(* IEC 61131-3 sources: traffic-lights/PLC_TrafficLights/Class/SafetyCDIAS_Base (part 5) *)

  // if there is a domain info attached
  if (pNameNewElement^ = '@') & ((pNameNewElement + 1)^ = 'D') then
    // check if it's in the actual domain
    if (pNameNewElement + 3)^ = ':' then
      // 1 digit domain number
      RemoteDomain := (pNameNewElement + 2)^ - '0';
    elsif (pNameNewElement + 4)^ = ':' then
      // 2 digits domain number
      RemoteDomain := ((pNameNewElement + 2)^ - '0') * 10 + (pNameNewElement + 3)^ - '0';
    else
      LogError("@ZZZZ (SafetyCDIAS_Base::AddUnsafeRoutElement) Invalid domain info at unsafe variable");
      return;
    end_if;

    // prepare the string (remove the domain info)
    if RemoteDomain >= 10 then
      ui_NameLen      -= 5;
      pNameNewElement += 5;
    else
      ui_NameLen      -= 4;
      pNameNewElement += 4;
    end_if;
  end_if;

  //With the first element, the table must be positioned
  if ( pRoutTable^ = NIL ) then

    //allocate memory for first routing element
    pRoutTable^$^void := To_StdLib.Malloc(size := sizeof(UnsafeIORoutingElement));

    if ( pRoutTable^ = NIL ) then

      State.uiIO_Flags                  := 0;
      State.uiIO_Flags.PhysicAccessOff 	:= 1;
      sd_retval                         :=-1;
      ClassState                        := _MemAllocFailed;
      return;

    end_if;

    p_RoutElement := pRoutTable^;

  else

    //add new element

    //add space for one element to table (linked list element for inputs and linear data area for outputs)
    if LinearMemory = FALSE then
    // search for a place
      p_RoutElement := pRoutTable^;
      while p_RoutElement^.pNext do
        p_RoutElement := p_RoutElement^.pNext;
      end_while;
      p_RoutElement^.pNext$^void := To_StdLib.Malloc(sizeof(UnsafeIORoutingElement));

      if ( p_RoutElement^.pNext = NIL ) then

        State.uiIO_Flags                  := 0;
        State.uiIO_Flags.PhysicAccessOff 	:= 1;
        sd_retval                         :=-1;
        ClassState                        := _MemAllocFailed;
        return;

      end_if;

      // set pointer to new element
      p_RoutElement := p_RoutElement^.pNext;
    else
      pRoutTable^$^void := To_StdLib.ReAlloc(mptr := pRoutTable^, newsize := ( ( pRoutElementsNo^ + 1 ) * sizeof(UnsafeIORoutingElement)));

      if ( pRoutTable^ = NIL ) then

        State.uiIO_Flags                  := 0;
        State.uiIO_Flags.PhysicAccessOff 	:= 1;
        sd_retval                         :=-1;
        ClassState                        := _MemAllocFailed;
        return;

      end_if;

      //set pointer to empty element on last position
      p_RoutElement := pRoutTable^ + ( pRoutElementsNo^ ) * sizeof(UnsafeIORoutingElement);
    end_if;
  end_if;

  if p_RoutElement then
    //allocate memory for name
    p_RoutElement^.pName$^void := To_StdLib.Malloc(size := ui_NameLen);

    if ( p_RoutElement^.pName = NIL ) then

      State.uiIO_Flags                  := 0;
      State.uiIO_Flags.PhysicAccessOff 	:= 1;
      sd_retval                         :=-1;
      ClassState                        := _MemAllocFailed;
      return;

    end_if;

    p_RoutElement^.NameLength := ui_NameLen;
    _memcpy(ptr1:=p_RoutElement^.pName, ptr2:=pNameNewElement, cntr:=ui_NameLen);

    // unsafe bdint variables are localized in a different memory area
    if BitMask then
      p_RoutElement^.ud_Address         := SDO_ADDRESS_UNSAFE_BDINT + ud_Address;
    else
      p_RoutElement^.ud_Address         := SDO_ADDRESS_APP_DATA + ud_Address;
    end_if;

    p_RoutElement^.BitMask              := BitMask;

    // initialize with invalid
    p_RoutElement^.b_IsValid            := FALSE;
    p_RoutElement^.sd_OldValue          := (16#80000000)$DINT;
    p_RoutElement^.sd_NewValue4External := (16#80000000)$DINT;

    // remember that we haven't transmitted this value so far
    p_RoutElement^.b_AlreadyTransmitted := FALSE;

    // initialize next pointer
    p_RoutElement^.pNext                := NIL;

    //increase counter
    pRoutElementsNo^                    += 1;

    // check if name exists in PLC
    p_RoutElement^.ud_Thisp             := GetThisViaServerName(pNameNewElement)$UDINT;
    if (pRoutTable = #p_UnsafeOutputsTable) & p_RoutElement^.BitMask then
      p_RoutElement^.UnsafeType         := BDINTOutput;
    else
      p_RoutElement^.UnsafeType         := NormalUnsafe;
    end_if;
  end_if;

END_FUNCTION

FUNCTION VIRTUAL SafetyCDIAS_Base::InitPathInfo
	VAR_INPUT
		pPathInfo 	: ^PathInfoType;
	END_VAR

  pPathInfo^.p_us_Path      := NIL;
  pPathInfo^.p_us_PathComp  := NIL;
  pPathInfo^.ui_PathCompLen := 0;

END_FUNCTION

FUNCTION VIRTUAL SafetyCDIAS_Base::WriteTDO2Module
	VAR_INPUT
		pTDO 	: ^TDOType;
	END_VAR
#ifdef SAFETY_OVER_DIAS
  VAR
    i : DINT;
  END_VAR
#endif

  if ( State.uiIO_Flags = 0 ) then

  #ifdef SAFETY_OVER_DIAS
    #pragma message("TDO-Handling over DIAS has to be reworked!")
    if ( b_im ) then
      //copy TDO word by word
      for i := 0 to (((TDOInfo AND 16#7F)/2)-1) by 1 do

        ( a_Handle_TDO_Write[i] )$^UINT^ := ( (pTDO)$^UINT + ( i * 2 ) )^;

      end_for;
    else
  #endif

      // responses into response buffer, request into requestbuffer (only enough place for 1)
      if pTDO^.StdHeader.Typ AND SSDO_MASK_RESPONSE then
        IF ( s_TDORingbuffer.ud_entries < ( SIZEOF( TDORingbuffer.Entry ) / SIZEOF( TDOType ) ) ) THEN
          s_TDORingbuffer.Entry[s_TDORingbuffer.ud_WritePos] :=  pTDO^;
          s_TDORingbuffer.ud_WritePos       := ( s_TDORingbuffer.ud_WritePos + 1 ) mod ( SIZEOF( TDORingbuffer.Entry ) / SIZEOF( TDOType ) );
          s_TDORingbuffer.ud_Entries        += 1;
          s_TDORingbuffer.b_ErrorTriggered  := FALSE;
        ELSIF ( s_TDORingbuffer.b_ErrorTriggered = FALSE ) THEN
          LogError("@ZZZZ (SafetyCDIAS_Base::WriteTDO2Module) [SL] Buffer for TDO-Messages is full!");
          s_TDORingbuffer.b_ErrorTriggered  := TRUE;
        END_IF;

        IF s_TDORingbuffer.ud_Entries > s_TDORingbuffer.ud_maxEntries THEN
          s_TDORingbuffer.ud_maxEntries     := s_TDORingbuffer.ud_Entries;
        END_IF;
      else
        s_TDORingbuffer.RequestTDO          := pTDO^;
        s_TDORingbuffer.b_RequestAvailable  := TRUE;
      end_if;

  #ifdef SAFETY_OVER_DIAS
    end_if;
  #endif
  end_if;

END_FUNCTION

FUNCTION VIRTUAL SafetyCDIAS_Base::ResetConfig
  VAR
    p_SafetyBase        : pVirtualBase;
  	p_RoutElement       : ^RoutElement;
    p_UnsafeRoutElement : ^UnsafeIORoutingElement;
    i                   : UINT;
    ii                  : DINT;
		MyPara 	            : CmdStruct;
		MyResult	          : results;
  END_VAR

  // tell all modules, which are connected to this cpu (through the old configuration) that they should delete the cpu from their routing table
  // must be more than 1, because 1st is always own entry
  if p_RoutTable & (ui_CntRoutElements > 1) then
    //set pointer on 2nd routing element
    p_RoutElement := p_RoutTable + sizeof(RoutElement);
    for i := 1 to (ui_CntRoutElements - 1) do
      // clear everything except this object (done after the for loop)
      if p_RoutElement^.ud_Thisp <> THIS$UDINT then
        // get thispointer of routing element
        p_SafetyBase := (p_RoutElement^.ud_Thisp)$pVirtualBase;

        // call other safety-class to remove the safetynumber from the routing table
        MyPara.uiCmd := CMD_SM_REMOVE_CPU_FROM_TABLE;
        MyPara.aPara[0] := SafetyNumber$DINT;

        p_SafetyBase^.NewInst(#MyPara, #MyResult);

//        p_SafetyBase^.RemoveCPUFromTable(ud_SafetyNr := SafetyNumber);
      end_if;

      // free memory of compressed path
      if p_RoutElement^.p_CompressedPath then
        To_StdLib.Free(mptr:=p_RoutElement^.p_CompressedPath);
      end_if;

      // set pointer on next routing element
      p_RoutElement += sizeof(RoutElement);
    end_for;

    // reduce local routing table to the cpu's own entry
    ui_CntRoutElements := 1;
  end_if;

  // on CSCP011 the SDO_COMMAND_WRITE_VALUES didn't exist, so we have to make a difference here
  if (us_Variant <> CSCP011_Preliminary) & (us_Variant <> CSCP011_Preliminary) then
    while p_UnsafeInputsTable do
      p_UnsafeRoutElement := p_UnsafeInputsTable;
      p_UnsafeInputsTable := p_UnsafeInputsTable^.pNext;

      To_StdLib.Free(mptr:=p_UnsafeRoutElement^.pName);
      To_StdLib.Free(mptr:=p_UnsafeRoutElement);
    end_while;
  else
    // free list of unsafe elements
    if p_UnsafeInputsTable then
      To_StdLib.Free(mptr:=p_UnsafeInputsTable);
      p_UnsafeInputsTable := NIL;
    end_if;
  end_if;
  ui_CntUnsafeInputs    := 0;

  // unsafe outputs are always in linear memory
  if p_UnsafeOutputsTable then
    To_StdLib.Free(mptr:=p_UnsafeOutputsTable);
    p_UnsafeOutputsTable := NIL;
  end_if;
  ui_CntUnsafeOutputs   := 0;

  // reset no of SDO input buffer
  ui_cnt_SDOInputBuffer := 0;

  // if the old configuration is reset, check for the configured state of the cpu
  b_CheckConfigured     := TRUE;

  if b_VaranAvailable then
    // by default the mover is invalid. it will be initialized when reading the configuration
    b_MoveCommandInputActive  := _Invalid;
    b_MoveCommandOutputActive := _Invalid;

    if b_PayloadSupport then

      DisableDO(ud_DOHandle := InputMovHandle$UDINT);

      if AdditionalSPDOs then
        for ii := 0 to (AdditionalSPDOs-1) do
          DisableDO(ud_DOHandle := aAdditionalPDOs[ii].InputMovHandle$UDINT);
        end_for;
      end_if;
    else

      if InputMovHandle then
        InputMovHandle^.ucCtrlStat := VARAN_DO_NO_RUN;
      end_if;

      if AdditionalSPDOs then
        for ii := 0 to (AdditionalSPDOs-1) do
          aAdditionalPDOs[ii].InputMovHandle^.ucCtrlStat := VARAN_DO_NO_RUN;
        end_for;
      end_if;
    end_if;

  else
    // if no VARAN, we can't move the PDOs
    b_MoveCommandInputActive  := _Inactive;
    b_MoveCommandOutputActive := _Inactive;
  end_if;

END_FUNCTION

FUNCTION VIRTUAL GLOBAL SafetyCDIAS_Base::MyBackground
  VAR
  	sd_retval         : DINT;
    GetStateResp      : GetStateResponseType;
    LastWriteCounter  : UDINT;
    FileHandle        : DINT;
		MyPara 	          : CmdStruct;
		MyResult	        : results;
  END_VAR

  // if any LED is active, then firmware update is not active and we can do our work
  if (VoltageOK | RunState | ServiceMode | Error) then

    // if a quit error is pending
    if QuitComError = 2 then
      MyPara.uiCmd := CMD_SM_QUIT_ERROR_VIA_OS;
      MyPara.aPara[0] := THIS$DINT;
      MyPara.aPara[1] := SafetyNumber$DINT;
      pSafetyManagerThis^.NewInst(#MyPara, #MyResult);

      QuitComError := MyResult.aData[0]$DINT;
    end_if;

    if (ClassState = _ReinitConfig) then

      // check every second if the cpu is configured
      if b_CheckConfigured & ((ops.tAbsolute - ud_LastCheckConfig) > 3000) then
        // get state via SDO communication
        sd_retval := SDOStdRequ ( us_Command      := SDO_COMMAND_GET_STATE
                                , p_us_RespData   := ( #GetStateResp )$^USINT
                                , us_RespLength   := sizeof(GetStateResponseType)
                                );

        // the cpu is configured, load the new configuration
        if ( sd_retval = 0 ) &
           (GetStateResp.ConfigState <> CFG_STATE_UNKNOWN) &
           (GetStateResp.ConfigState <> CFG_STATE_INVALID) &
           (GetStateResp.ConfigState <> CFG_STATE_NOT_CONFIGURED) then

          b_CheckConfigured := FALSE;
          b_GetNewConfiguration := TRUE;
        end_if;

        // remember the last time we checked for configurated cpu
        ud_LastCheckConfig := ops.tAbsolute;
      end_if;

      // if there is a new configuration => get it
      if b_GetNewConfiguration then

        //get configuration from safe CPU and build routing tables
        sd_retval := GetRoutingData();
        if sd_retval = 0 then
          b_GetNewConfiguration := FALSE;

          SendAllUnsafeValues();
        else
          LogError("@ZZZZ (SafetyCDIAS_Base::MyBackground) FAILED TO REINIT THE SAFECPU: ");
        end_if;
      end_if;
    end_if;

    // here we save the log file from the module to the harddrive (started by user)
    if DiagVars.SavingLogInProgress then

      case DiagVars.SavingLogSSW of

  // ********************************************************************************************************************************************
        GetLogHeader:     // get log header from module (contains size of log memory and write counter)

          // get log header via SDO communication
          sd_retval := SDORequ ( us_Command      := SDO_COMMAND_GET_LOG_HDR
                               , p_us_RequData   := #DiagVars.ucChoiceSaveLog
                               , us_RequLength   := 1
                               , p_us_RespData   := ( #DiagVars.LogHeader)$^USINT
                               , us_RespLength   := sizeof(DiagStructType.LogHeader)
                               );

          if ( sd_retval = 0 ) then
            DiagVars.LogMemToGet := DiagVars.LogHeader.LogMemSize;
            DiagVars.pLogFileMem$pVoid := To_StdLib.Malloc(size:=DiagVars.LogHeader.LogMemSize);
            //_memset(dest:=DiagVars.pLogFileMem$pVoid, usByte:=0, cntr:=DiagVars.LogHeader.LogMemSize);
            if DiagVars.ucChoiceSaveLog = 0 then
              DiagVars.ReadBaseAdr  := SDO_ADDRESS_LOG_UC1;
            else
              DiagVars.ReadBaseAdr  := SDO_ADDRESS_LOG_UC2;
            end_if;
            DiagVars.SavingLogSSW   := GetLogFileBlocks;

          end_if;

  // ********************************************************************************************************************************************
        GetLogFileBlocks: // get the log memory from the application memory of the module (every cycle only a little bit to prevent runtime error in module)

          // we wait here until UpdateCy finishes our work

  // ********************************************************************************************************************************************
        GetLogHeader2:    // get log header from module again. if write counter changed,
                          // we repeat GetLogFileBlocks. otherwise we continue to save the file

          LastWriteCounter := DiagVars.LogHeader.WriteCounter;

          // get LogHeader
          sd_retval := SDORequ ( us_Command      := SDO_COMMAND_GET_LOG_HDR
                               , p_us_RequData   := #DiagVars.ucChoiceSaveLog
                               , us_RequLength   := 1
                               , p_us_RespData   := ( #DiagVars.LogHeader)$^USINT
                               , us_RespLength   := sizeof(DiagStructType.LogHeader)
                               );

          if ( sd_retval = 0 ) then

            // if write counter is different, repeat last step
            if DiagVars.LogHeader.WriteCounter <> LastWriteCounter then
              DiagVars.SavingLogSSW := GetLogFileBlocks;

              DiagVars.LogMemToGet := DiagVars.LogHeader.LogMemSize;

              // realloc memory (maybe it's a different size)
              To_StdLib.Free(mptr:=DiagVars.pLogFileMem$pVoid);
              DiagVars.pLogFileMem$pVoid := To_StdLib.Malloc(size:=DiagVars.LogHeader.LogMemSize);
            else
              // write counter is equal. continue to last step
              DiagVars.SavingLogSSW := SaveLogFile;
            end_if;
          end_if;

  // ********************************************************************************************************************************************
        SaveLogFile:      // save the memory to the specified file (DPNE)
          // open file (create/overwrite always)
          FileHandle := FileSys.FileOpen(filename:=#DiagVars.DPNE[0], attributes:=ATT_CREATE_ALWAYS);

          DiagVars.SavingLogSuccessful := 1;

          if FileHandle >= 0 then

            // save content to it
            if FileSys.FileWrite(handle:=FileHandle, buffer:=DiagVars.pLogFileMem, length:=DiagVars.LogHeader.LogMemSize) <> DiagVars.LogHeader.LogMemSize$DINT then
              // failed to write to file
              LogError("@ZZZZ (SafetyCDIAS_Base::MyBackground) Failed to write to binary LogFile");
              DiagVars.SavingLogSuccessful := -1;
            end_if;

            // close file
            FileSys.FileClose(handle:=FileHandle);
          else
            // failed to open file
            LogError("@ZZZZ (SafetyCDIAS_Base::MyBackground) Failed to open binary LogFile");
            DiagVars.SavingLogSuccessful := -1;
          end_if;

          To_StdLib.Free(mptr:=DiagVars.pLogFileMem$pVoid);
          DiagVars.pLogFileMem := NIL;

          DiagVars.SavingLogSSW         := GetLogHeader;
          DiagVars.SavingLogInProgress  := FALSE;

      end_case;
    end_if;
  end_if;

END_FUNCTION

FUNCTION VIRTUAL SafetyCDIAS_Base::RemoveCPUFromTable
	VAR_INPUT
		ud_SafetyNr 	  : HDINT;
	END_VAR
  VAR
  	p_RoutElement   : ^RoutElement;
    i               : UDINT;
    FoundIndex      : UDINT;
    pPDOInputBuffer : ^PDOInputBuffer;
    Found : BOOL;
  END_VAR

  // if we are a cpu, do nothing
  if b_CheckCRC then
    return;
  end_if;

  //check each element (must be more than 1, because 1st is always own entry)
  if p_RoutTable & (ui_CntRoutElements > 1) then
    //set pointer on 2nd routing element
    p_RoutElement := p_RoutTable + sizeof(RoutElement);
    for i := 1 to (ui_CntRoutElements - 1) do

      // if we found safenumber, delete element from table
      if ( p_RoutElement^.ud_SafeNumber = ud_SafetyNr ) then

        // at last element we don't need to copy data, just decrease buffersize
        if i <> (ui_CntRoutElements - 1) then
          _memcpy(p_RoutElement, p_RoutElement + sizeof(RoutElement), sizeof(RoutElement) * (ui_CntRoutElements - 1 - i));
        end_if;

        // free 1 element and decrease element counter
        ui_CntRoutElements -= 1;

        exit;
      end_if;

      // set pointer on next routing element
      p_RoutElement += sizeof(RoutElement);
    end_for;
  end_if;

  // reset no of SDO input buffer
  ui_cnt_SDOInputBuffer := 0;

  if b_VaranAvailable then
    // by default the mover is invalid. it will be initialized when reading the configuration
    b_MoveCommandInputActive  := _Invalid;
    b_MoveCommandOutputActive := _Invalid;

    if InputMovHandle then
      if b_PayloadSupport then
        DisableDO(ud_DOHandle := InputMovHandle$UDINT);

        if AdditionalSPDOs then
          for i := 0 to (AdditionalSPDOs-1)$UDINT do
            DisableDO(ud_DOHandle := aAdditionalPDOs[i].InputMovHandle$UDINT);
          end_for;
        end_if;
      else
        InputMovHandle^.ucCtrlStat := VARAN_DO_NO_RUN;

        if AdditionalSPDOs then
          for i := 0 to (AdditionalSPDOs-1)$UDINT do
            aAdditionalPDOs[i].InputMovHandle^.ucCtrlStat := VARAN_DO_NO_RUN;
          end_for;
        end_if;

      end_if;
    end_if;
  else
    // if no VARAN, we can't move the PDOs
    b_MoveCommandInputActive  := _Inactive;
    b_MoveCommandOutputActive := _Inactive;
  end_if;

  // check if we received a PDO from this CPU => if so, delete it from the PDO input buffer
  if ui_cnt_PDOInputBuffer then
    // search for the PDO
    Found := FALSE;
    pPDOInputBuffer := #aPDOInputBuffer[0];
    for FoundIndex := 0 to (ui_cnt_PDOInputBuffer-1) do
      if pPDOInputBuffer^.ud_SafetyNr = ud_SafetyNr then
        Found := TRUE;
        exit;
      end_if;

      pPDOInputBuffer += sizeof(PDOInputBuffer);
    end_for;

    // if we found the PDO => remove it from memory (move the memory behind the found PDO over the place of the found PDO)
    if Found then
      // if it's last entry (no entries have to be moved) => we only have to copy some memory if it's not the last
      if FoundIndex < (ui_cnt_PDOInputBuffer-1) then
        for i := FoundIndex to (ui_cnt_PDOInputBuffer-2) do
          aPDOInputBuffer[i] := aPDOInputBuffer[i+1];
        end_for;
      end_if;
      ui_cnt_PDOInputBuffer -= 1;
    end_if;
  end_if;

END_FUNCTION

FUNCTION VIRTUAL SafetyCDIAS_Base::CheckUnsafeUpdateCycle

  // we can only use 56 byte pay load (instead of 64) because fw drops the 8 byte used for addresses in safe SDO

  if ui_CntUnsafeOutputs then
  // maximum of read variables in 1 frame is 15 (56 Bytes pay load - 1 Byte Returncode - 1 Byte Length = 54 Bytes => 13x4Bytes = 52)
    MaxVarsPerReadPackage := (SDO_MAX_LENGTH - (sizeof(SDOHeader) - sizeof(SDOHeader.SessId)) - sizeof(SDORespReadConfig.us_Returncode) - sizeof(SDORespReadConfig.us_Length)) / sizeof(DINT);
    ReadFramesNeeded := ((ui_CntUnsafeOutputs - 1) / MaxVarsPerReadPackage) + 1;
  else
    ReadFramesNeeded := 0;
  end_if;

  if ui_CntUnsafeInputs then
  // maximum of write variables in 1 frame is 14 (56 Bytes pay load - 4 Byte Address - 1 Byte Length = 51 Bytes => 12x4Bytes = 48)
    MaxVarsPerWritePackage := (SDO_MAX_LENGTH - (sizeof(SDOHeader) - sizeof(SDOHeader.SessId)) - sizeof(SDORequReadConfig.ud_Address) - sizeof(SDORequReadConfig.us_Length)) / sizeof(DINT);
    WriteFramesNeeded := ((ui_CntUnsafeInputs - 1) / MaxVarsPerWritePackage) + 1;
  else
    WriteFramesNeeded := 0;
  end_if;

  // check if user has given us enough time
  if b_VaranAvailable then
    if sd_VaranType = 2 then
      ud_TransfertimePerPackage := SDO_TRANSFERTIME_MOVER;
    else
      ud_TransfertimePerPackage := SDO_TRANSFERTIME_VARAN;
    end_if;
  else
    ud_TransfertimePerPackage := SDO_TRANSFERTIME_CDIAS;
#ifdef SAFETY_OVER_DIAS
    #pragma message("Transfer time for DIAS must be defined!")
#endif
  end_if;

  if ( (WriteFramesNeeded + ReadFramesNeeded) * ud_TransfertimePerPackage ) > ServerUpdateTime then
    ServerUpdateTime    := ( WriteFramesNeeded + ReadFramesNeeded ) * ud_TransfertimePerPackage;
    ServerUpdateTime.Write(input:=ServerUpdateTime);
    ud_ServerUpdateTime := ( ReadFramesNeeded ) * ud_TransfertimePerPackage;
  end_if;

END_FUNCTION

FUNCTION VIRTUAL GLOBAL SafetyCDIAS_Base::FetchDiagState

  DiagVars.UserDiagStateReady := FALSE;
  DiagVars.UserWantsDiagState := TRUE;

END_FUNCTION

FUNCTION VIRTUAL GLOBAL SafetyCDIAS_Base::GetDiagState
	VAR_INPUT
		pDiagState 	: ^SafetyDiagState;
	END_VAR
	VAR_OUTPUT
		StateReady 	: BOOL;
	END_VAR

  StateReady                        := DiagVars.UserDiagStateReady;

  // if data ready, we save it into user structure
  if StateReady then
    pDiagState^.RunState            := DiagVars.UserGetStateResp.RuntimeState;
    pDiagState^.ConfigState         := DiagVars.UserGetStateResp.ConfigState;
    pDiagState^.LoginLevel          := DiagVars.UserGetStateResp.LoginLevel;
    pDiagState^.ErrorCounterIOState := DiagVars.UserGetStateResp.ErrorCount;
  end_if;

END_FUNCTION

FUNCTION VIRTUAL GLOBAL SafetyCDIAS_Base::FetchDiagInfo
	VAR_INPUT
		ucChoice 	: USINT;
	END_VAR

  DiagVars.ucChoiceDiagInfo  := ucChoice;
  DiagVars.UserDiagInfoReady := FALSE;
  DiagVars.UserWantsDiagInfo := TRUE;

END_FUNCTION

FUNCTION VIRTUAL GLOBAL SafetyCDIAS_Base::GetDiagInfo
	VAR_INPUT
		pDiagInfo 	: ^SafetyDiagInfo;
	END_VAR
	VAR_OUTPUT
		StateReady 	: BOOL;
	END_VAR

  StateReady    := DiagVars.UserDiagInfoReady;

  // if data ready, we save it into user structure
  if StateReady then
    pDiagInfo^  := DiagVars.UserGetDiagInfoResp;
  end_if;

END_FUNCTION

FUNCTION VIRTUAL SafetyCDIAS_Base::SDORequ
	VAR_INPUT
		us_Command 	        : USINT;
		p_us_RequData 	    : ^USINT;
		us_RequLength 	    : USINT;
		p_us_RespData 	    : ^USINT;
		us_RespLength 	    : USINT;
	END_VAR
	VAR_OUTPUT
		sd_retval 	        : DINT;
	END_VAR
  VAR
  	pSDORequestBuffer   : ^SDOStdHeader;
    pSDOResponseBuffer  : ^SDOStdResp;
    RespBuffer          : ARRAY [0..127] OF USINT;
    RequBuffer          : ARRAY [0..127] OF USINT;
    us_InLength         : USINT;
    us_OutLength        : USINT;
  END_VAR

  //SDO requests for this commands don't have any further data
  pSDORequestBuffer$^void   := #RequBuffer[0];
  pSDOResponseBuffer$^void  := #RespBuffer[0];

  //SDO request buffer (length header + data)
  us_InLength               := sizeof(SDOStdHeader) + us_RequLength;

  //SDO response buffer (length header + rc + data)
  us_OutLength              := sizeof(SDOStdHeader) + 1 + us_RespLength;

  //calculate length without crc
  pSDORequestBuffer^.len    := sizeof(SDOStdHeader) - sizeof(SDOStdHeader.CRC) + us_RequLength;

  //type
  pSDORequestBuffer^.typ    := FRM_TYPECODE_STD;

  //sequence number
  pSDORequestBuffer^.SeqNr  := us_CntSequNr;

  _memcpy(ptr1:=pSDORequestBuffer + sizeof(SDOStdHeader), ptr2:=p_us_RequData, cntr:=us_RequLength);

  //increase counter for sequence number
  if us_CntSequNr < 16#7F then
    us_CntSequNr += 1;
  else
    us_CntSequNr := 0;
  end_if;

  //command to inform CPU about initializing classes is ok
  pSDORequestBuffer^.cmd := us_Command;

  //set CRC-field to 0
  pSDORequestBuffer^.CRC := 0;

  //send request
  sd_retval := SAFETY_iSendRequest( uiMaster    := 0
                                  , pucNode     := p_ObjectPath
                                  , uiInLength  := us_InLength
                                  , pucInput    := pSDORequestBuffer$^USINT
                                  , uiOutLength := us_OutLength
                                  , pucOutput   := pSDOResponseBuffer$^USINT
                                  );

  //no response
  if ( sd_retval = 0 ) then

    //check sequence number to exclude a possible wrong response
    if ( pSDORequestBuffer^.SeqNr <> pSDOResponseBuffer^.StdHeader.SeqNr ) then
      sd_retval := -102;

    //check returncode of SDO
    elsif ( pSDOResponseBuffer^.us_Returncode <> SDO_RETCODE_OK ) then
      sd_retval := -103;
    end_if;

  end_if;

  //return response
  if ( ( sd_retval = 0 ) & ( p_us_RespData <> NIL )) then
    To_StdLib.MemCpy(dest := p_us_RespData, source := #pSDOResponseBuffer^.us_Data, size := us_RespLength);
  end_if;

END_FUNCTION

FUNCTION VIRTUAL GLOBAL SafetyCDIAS_Base::SaveLog
	VAR_INPUT
		ucChoice  : USINT;
		pDPNE 	  : ^CHAR;
	END_VAR
	VAR_OUTPUT
		Success 	: DINT;
	END_VAR

  if DiagVars.SavingLogInProgress = FALSE then
    DiagVars.SavingLogInProgress  := TRUE;

    DiagVars.SavingLogSuccessful  := FALSE; //Reset Value

    DiagVars.ucChoiceSaveLog      := ucChoice;

    _memcpy(ptr1:=#DiagVars.DPNE, ptr2:=pDPNE, cntr:=_strlen(pDPNE));

    Success := TRUE;
  else
    Success := FALSE;
  end_if;

END_FUNCTION

FUNCTION VIRTUAL GLOBAL SafetyCDIAS_Base::SaveLogActive
	VAR_OUTPUT
		InProgress 	: BOOL;
	END_VAR

  InProgress := DiagVars.SavingLogInProgress;

END_FUNCTION

FUNCTION VIRTUAL SafetyCDIAS_Base::BlockedTransferLength
	VAR_INPUT
		ud_Datalength 	    : UDINT;
		us_MaxBlocklength 	: USINT;
	END_VAR
	VAR_OUTPUT
		us_ActBlocklength 	: USINT;
	END_VAR

  IF ud_Datalength > to_UDINT(us_MaxBlocklength) THEN
    us_ActBlocklength := us_MaxBlocklength;
  ELSE
    us_ActBlocklength := to_USINT(ud_Datalength);
  END_IF;

END_FUNCTION

FUNCTION VIRTUAL SafetyCDIAS_Base::AddToPDOMoverList
	VAR_INPUT
		pThis 	: pVirtualBase;
		pList 	: ^pPDOMoverList;
	END_VAR
  VAR
    pHelp : ^PDOMoverList;
  END_VAR

  if pList^ = NIL then
    pList$^pvoid^ := To_StdLib.Malloc(size:=sizeof(PDOMoverList));
    //Graphic.Memory((#pList)$^pVoid, sizeof(PDOMoverList));
    pHelp := pList^;
  else
    pHelp := pList^;
    if pHelp^.pThis = pThis then
      // this pointer already in buffer => leave function
      return;
    end_if;
    while pHelp^.pNext <> NIL do
      if pHelp^.pThis <> pThis then
        pHelp := pHelp^.pNext;
      else
        // this pointer already in buffer => leave function
        return;
      end_if;
    end_while;
    pHelp^.pNext$pvoid := To_StdLib.Malloc(size:=sizeof(PDOMoverList));
    pHelp := pHelp^.pNext;
  end_if;

  if pHelp <> NIL then
    pHelp^.pThis := pThis;
    pHelp^.pNext := NIL;
  end_if;

END_FUNCTION

FUNCTION VIRTUAL SafetyCDIAS_Base::WalkThroughPDOMoverList
	VAR_INPUT
		pList 	  : ^pPDOMoverList;
		NewState 	: PDOMoveState;
	END_VAR
  VAR
  	pAct      : ^PDOMoverList;
    pFree     : ^void;
		MyPara 	  : CmdStruct;
		MyResult  : results;
  END_VAR

  // get pointer on first element of list
  pAct := pList^;

  // if we have entries left we walk on
  WHILE pAct DO
#pragma warning(disable:137 )
    // set state of corresponding PDOMover to off
    IF pList = #pPDOMoverListInputs THEN
      if NewState = _Inactive then

        MyPara.uiCmd    := CMD_SM_DEACTIVATE_MOVE_CMD;
        MyPara.aPara[0] := 0;
        pAct^.pThis^.NewInst(#MyPara, #MyResult);

//        pAct^.pThis^.b_MoveCommandOutputActive := _Inactive;
      end_if;
    ELSE
      if NewState = _Inactive then

        MyPara.uiCmd    := CMD_SM_DEACTIVATE_MOVE_CMD;
        MyPara.aPara[0] := 1;
        pAct^.pThis^.NewInst(#MyPara, #MyResult);

//        pAct^.pThis^.b_MoveCommandInputActive := _Inactive;
      end_if;
    END_IF;
#pragma warning(default:137 )

    //go to next entry and get rid of the allocated memory
    pFree := pAct;
    pAct  := pAct^.pNext;
    To_StdLib.Free(mptr:=pFree);
  END_WHILE;

  // we got rid of the memory above - to make sure nobody will use this data again we clear the list entry
  pList^ := NIL;

END_FUNCTION

FUNCTION VIRTUAL SafetyCDIAS_Base::CleanupPDOMoverList
	VAR_INPUT
		pList 	: ^pPDOMoverList;
	END_VAR
  VAR
  	pAct    : ^PDOMoverList;
    pFree   : ^void;
  END_VAR

  // get pointer on first element of list
  pAct := pList^;

  // if we have entries left we walk on
  WHILE pAct DO
    //go to next entry and get rid of the allocated memory
    pFree := pAct;
    pAct  := pAct^.pNext;
    To_StdLib.Free(mptr:=pFree);
  END_WHILE;

  // we got rid of the memory above - to make sure nobody will use this data again we clear the list entry
  pList^ := NIL;

END_FUNCTION

#pragma warning(disable: 73)
FUNCTION VIRTUAL SafetyCDIAS_Base::AddFrame
	VAR_INPUT
		pFrame 	        : ^SafetyCDIAS_Base::SDOStdHeader;
		FrameState 	    : DINT;
		CallerSafetyNr 	: HDINT;
	END_VAR

END_FUNCTION
#pragma warning(default: 73)

FUNCTION VIRTUAL SafetyCDIAS_Base::RecordFrame
	VAR_INPUT
		pFrame 	    : ^DINT;
		FrameState 	: DINT;
	END_VAR
  VAR
    ThisBackup  : pVoid;
    TempSafetyNr: HDINT;
  END_VAR

  if pAnalyzerThis & pAnalyzerMethod then

    TempSafetyNr  := SafetyNumber;

    ThisBackup    := THIS;

    THIS          := pAnalyzerThis$^SafetyCDIAS_Base;
    pAnalyzerMethod$AddFrame(pFrame$^SDOStdHeader, FrameState, TempSafetyNr);

    THIS          := ThisBackup$^SafetyCDIAS_Base;
  end_if;

END_FUNCTION

#pragma warning(disable: 73)
FUNCTION VIRTUAL GLOBAL SafetyCDIAS_Base::UpDateRTPostScan
	VAR_INPUT
		Handle 	          : UDINT;
	END_VAR
  VAR
  	i                 : UDINT;
    TempSafetyNr      : HDINT;
    p_PDOInBufferAct  : ^PDOInputBuffer;
  END_VAR

//============================ Profiler start======================================================
#ifdef  DM_Profiler
  StartTimeMeasurement(usMode := DMTIME_RTPOSTSCAN);
#endif
//============================ Profiler end========================================================

  // do tdo/pdo communication only, if module has been found and initialized correctly and if there are some LEDs on (else a FW-Update is running)
  if ( State.uiIO_Flags = 0 ) &
     (( ClassState = _SafetyClassOK ) | ( ClassState = _WaitForSynchronicity ) | ( ClassState = _ModFromCfgNotFound ) | ( ClassState = _UnknownCfgError ) | ( ClassState = _UnsafeVarNotFound )) then

    // if any LED is active, then firmware update is not active and we can do our work
    if (VoltageOK | RunState | ServiceMode | Error) then

      // write unsafe I/Os
      UpDateNotStd(calloption:=CALL_OPTION_RT_POSTSCAN);

      // TDO Handling with mover
      if TDOSingleRunActive then
        TDOSingleRunActive := FALSE;
        if b_PayloadSupport then
          p_HandleTDOWriteEnable^     := VARAN_DO_NO_RUN;
        else
          ( p_HandleTDOWrite$^USINT )^  := VARAN_DO_NO_RUN;
        end_if;
      end_if;

      // check if we may send a TDO (TDO-Status-Register MSB must be zero)
      if (( p_us_Handle_TDO_Status_Write^ AND 16#80 ) = 0) then

        // check for a TDO Request => if there is one, send it
        if s_TDORingbuffer.b_RequestAvailable then

          To_StdLib.MemCpy(dest := p_us_Handle_TDO_Write, source := #s_TDORingbuffer.RequestTDO, size := sizeof(TDOType));

          TimeSyncDOActive.Wait4ResponseNo += 1;
#ifdef DO_DEBUG
          DOCheck(pFrame:=(#s_TDORingbuffer.RequestTDO)$^SDOStdHeader, pCheckStruct:=#TDOWrite);
#endif

#ifdef SAFETY_PROTOCOL_ANALYZER_ACTIVATED
  RecordFrame((#s_TDORingbuffer.RequestTDO)$^DINT, 1);
#endif

          s_TDORingbuffer.b_RequestAvailable := FALSE;

          if b_VaranAvailable then
            if (sd_VaranType = 1) then

              if b_PayloadSupport then  // Payload, No Mover ---------------------------------------------------------------------

                if b_DOIsRunningTDOWrite.StartRequest then  // Check if the startrequest has been set somewhere else, probably not the same check as without payload.
                  TDOErrorDetectedCnt += 1;
                end_if;

                b_DOIsRunningTDOWrite.StartRequest := true;

                if b_NewSyncMode then
                  // start DO at this point to ensure 1 cycle delay, from request to response
                  EnableDO(ud_DOHandle := p_HandleTDORead$UDINT);
                  b_DOIsRunningTDORead.ContRun := true; // Important! This flag is checked in UpdataRT
                end_if;

              else  // No Payload, No Mover -------------------------------------------------------------------------------------------

                if p_HandleTDOWrite^.ucCtrlStat AND VARAN_DO_SINGLE_RUN then
                  TDOErrorDetectedCnt += 1;
                end_if;

                p_HandleTDOWrite^.ucCtrlStat  := VARAN_DO_SINGLE_RUN;

                if b_NewSyncMode then
                  // start DO at this point to ensure 1 cycle delay, from request to response
                  p_HandleTDORead^.ucCtrlStat := VARAN_DO_CONT_RUN;
                end_if;

              end_if;

            else  // Mover

              if b_PayloadSupport then  // Payload, Mover ---------------------------------------------------------------------

                if p_HandleTDOWriteEnable^ AND VARAN_MOVER_DO_SINGLE_RUN then
                  TDOErrorDetectedCnt += 1;
                end_if;
                  p_HandleTDOWriteEnable^ := VARAN_MOVER_DO_SINGLE_RUN;
                TDOSingleRunActive := TRUE;

              else  // No Payload, Mover -------------------------------------------------------------------------------------------

                if ( p_HandleTDOWrite$^USINT )^ AND VARAN_MOVER_DO_SINGLE_RUN then
                  TDOErrorDetectedCnt += 1;
                end_if;
                ( p_HandleTDOWrite$^USINT )^ := VARAN_MOVER_DO_SINGLE_RUN;
                TDOSingleRunActive := TRUE;

              end_if;
            end_if;
          end_if;

        // Send entries of TDO-Buffer (only responses)
        elsif ( s_TDORingbuffer.ud_Entries > 0 ) THEN

          To_StdLib.MemCpy(dest := p_us_Handle_TDO_Write, source := #s_TDORingbuffer.Entry[s_TDORingbuffer.ud_ReadPos], size := sizeof(TDOType));

#ifdef DO_DEBUG
          DOCheck(pFrame:=(#s_TDORingbuffer.Entry[s_TDORingbuffer.ud_ReadPos])$^SDOStdHeader, pCheckStruct:=#TDOWrite);
#endif

#ifdef SAFETY_PROTOCOL_ANALYZER_ACTIVATED
  RecordFrame((#s_TDORingbuffer.Entry[s_TDORingbuffer.ud_ReadPos])$^DINT, 1);
#endif

          // in the startupphase we use the time synchronisation between modules to check if a module is synchron with all of his communication partners
          if (us_SetBusReadyState = WaitPDOsSyncron) & ui_cnt_PDOInputBuffer then
            TempSafetyNr := s_TDORingbuffer.Entry[s_TDORingbuffer.ud_ReadPos].SrcAdr;

            p_PDOInBufferAct := #aPDOInputBuffer[0];
            for i := 0 to (ui_cnt_PDOInputBuffer-1) do
              if p_PDOInBufferAct^.ud_SafetyNr = TempSafetyNr then
                p_PDOInBufferAct^.b_TimeSynchron := TRUE;
              end_if;

              p_PDOInBufferAct +=  sizeof(PDOInputBuffer);
            end_for;
          end_if;

          s_TDORingbuffer.ud_ReadPos := ( s_TDORingbuffer.ud_ReadPos + 1 ) mod ( SIZEOF( TDORingbuffer.Entry ) / SIZEOF( TDOType ) );
          s_TDORingbuffer.ud_Entries -= 1;

          if b_VaranAvailable then
            if (sd_VaranType = 1) then

              if b_PayloadSupport then   // Payload, No Mover ---------------------------------------------------------------------
                if b_DOIsRunningTDOWrite.StartRequest then // Check if the startrequest has been set somewhere else, probably not the same check as without payload.
                  TDOErrorDetectedCnt += 1;
                end_if;

                b_DOIsRunningTDOWrite.StartRequest := true;

                if b_NewSyncMode then
                  // start DO at this point to ensure 1 cycle delay, from request to response
                  EnableDO(ud_DOHandle := p_HandleTDORead$UDINT);
                  b_DOIsRunningTDORead.ContRun := true; // Important! This flag is checked in UpdataRT
                end_if;

              else  // No Payload, No Mover -------------------------------------------------------------------------------------------

                if p_HandleTDOWrite^.ucCtrlStat AND VARAN_DO_SINGLE_RUN then
                  TDOErrorDetectedCnt += 1;
                end_if;

                p_HandleTDOWrite^.ucCtrlStat  := VARAN_DO_SINGLE_RUN;

                if b_NewSyncMode then
                  // start DO at this point to ensure 1 cycle delay, from request to response
                  p_HandleTDORead^.ucCtrlStat := VARAN_DO_CONT_RUN;
                end_if;

              end_if;

            else  // Mover

              if b_PayloadSupport then  // Payload, Mover ---------------------------------------------------------------------

                if p_HandleTDOWriteEnable^ AND VARAN_MOVER_DO_SINGLE_RUN then
                  TDOErrorDetectedCnt += 1;
                end_if;
                p_HandleTDOWriteEnable^ := VARAN_MOVER_DO_SINGLE_RUN;
                TDOSingleRunActive := TRUE;

              else  // No Payload, Mover -------------------------------------------------------------------------------------------

                if ( p_HandleTDOWrite$^USINT )^ AND VARAN_MOVER_DO_SINGLE_RUN then
                  TDOErrorDetectedCnt += 1;
                end_if;
                ( p_HandleTDOWrite$^USINT )^ := VARAN_MOVER_DO_SINGLE_RUN;
                TDOSingleRunActive := TRUE;

              end_if;

            end_if;
          end_if;
        END_IF;
      else
        // can't write this time, if there is a request waiting => drop it
        if s_TDORingbuffer.b_RequestAvailable then
          s_TDORingbuffer.b_RequestAvailable := FALSE;
          RequestDropCounter += 1;
        end_if;
      end_if;

      if RunState & ((us_SetBusReadyState = SetBusReadyFinished) | b_ManualQuit) then
        //write PDO to hardware
        if ( ui_cnt_PDOInputBuffer > 0 ) then
          WritePDO2Module();
        end_if;
      end_if;
    end_if;
  end_if;

  if b_PayloadSupport & (sd_VaranType = 1) then

    // p_HandleTDORead xxxxxxxxxxxxxxxxxxxxxxxxxxxxxxxxxxxxxxxxxxxxxxxxxxxxxxxxxxxxxxxxxxxxxxxxxxxxxxxxxxxxxxxxxxxxxxxx
    case b_DOIsRunningTDORead of

      SR_STATE_ENABLE_ME :  // DO is not running and start request is set ----------------------------------------
        EnableDO(ud_DOHandle  := p_HandleTDORead$UDINT);
        b_DOIsRunningTDORead  := SR_STATE_DISABLE_ME;

      SR_STATE_DISABLE_ME : // DO is running and start request is not set ----------------------------------------
        DisableDO(ud_DOHandle := p_HandleTDORead$UDINT);
        b_DOIsRunningTDORead  := SR_STATE_NOTHING;

      SR_STATE_LEAVE_ME_ENABLED : // DO is running and another start request is set ------------------------------
        b_DOIsRunningTDORead  := SR_STATE_DISABLE_ME;

    end_case;

    // p_HandleTDOWrite xxxxxxxxxxxxxxxxxxxxxxxxxxxxxxxxxxxxxxxxxxxxxxxxxxxxxxxxxxxxxxxxxxxxxxxxxxxxxxxxxxxxxxxxxxxxxxxx
    case b_DOIsRunningTDOWrite of

      SR_STATE_ENABLE_ME :  // DO is not running and start request is set ----------------------------------------
        EnableDO(ud_DOHandle  := p_HandleTDOWrite$UDINT);
        b_DOIsRunningTDOWrite := SR_STATE_DISABLE_ME;

      SR_STATE_DISABLE_ME : // DO is running and start request is not set ----------------------------------------
        DisableDO(ud_DOHandle := p_HandleTDOWrite$UDINT);
        b_DOIsRunningTDOWrite := SR_STATE_NOTHING;

      SR_STATE_LEAVE_ME_ENABLED : // DO is running and another start request is set ------------------------------
        b_DOIsRunningTDOWrite := SR_STATE_DISABLE_ME;

    end_case;

    // p_HandleUnsafeOutWrite xxxxxxxxxxxxxxxxxxxxxxxxxxxxxxxxxxxxxxxxxxxxxxxxxxxxxxxxxxxxxxxxxxxxxxxxxxxxxxxxxxxxxxxxxxxxxxxx
    case b_DOIsRunningUnsafeOutWrite of

      SR_STATE_ENABLE_ME :  // DO is not running and start request is set ----------------------------------------
        EnableDO(ud_DOHandle  := p_HandleUnsafeOutWrite$UDINT);
        b_DOIsRunningUnsafeOutWrite := SR_STATE_DISABLE_ME;

      SR_STATE_DISABLE_ME : // DO is running and start request is not set ----------------------------------------
        DisableDO(ud_DOHandle := p_HandleUnsafeOutWrite$UDINT);
        b_DOIsRunningUnsafeOutWrite := SR_STATE_NOTHING;

      SR_STATE_LEAVE_ME_ENABLED : // DO is running and another start request is set ------------------------------
        b_DOIsRunningUnsafeOutWrite := SR_STATE_DISABLE_ME;

    end_case;

  end_if;

//============================ Profiler start======================================================
#ifdef  DM_Profiler
  StopTimeMeasurement(usMode := DMTIME_RTPOSTSCAN);
#endif
//============================ Profiler end========================================================

END_FUNCTION
#pragma warning(default: 73)

FUNCTION VIRTUAL GLOBAL SafetyCDIAS_Base::State::NewInst
	VAR_INPUT
		pPara 	        : ^CmdStruct;
		pResult 	      : ^Results;
	END_VAR
	VAR_OUTPUT
		ret_code 	      : IprStates;
	END_VAR
  VAR
  	OldClassState   : SafetyConfigStateType;
    pPDOInputBuffer : ^PDOInputBuffer;
    i, j            : UINT;
    Found           : BOOL;
    sd_retval       : DINT;
    GetStateResp    : GetStateResponseType;

  	ptmpStr         : ^CHAR;
    ud_StrSize      : UDINT;
    us_temp         : USINT;

  END_VAR

	ret_code := READY;

	CASE pPara^.uiCmd OF
//**********************************************************************************************************************************************************
		CMD_SM_SET_NEW_SYNC_MODE:

      b_NewSyncMode := pPara^.aPara[0]$BOOL; //TRUE;

      if b_NewSyncMode then
        NewHandShakeValue := 2#001;
      end_if;

//**********************************************************************************************************************************************************
    CMD_SM_START_TIME_SYNC:

      // set bit for starting timesync at the module (bit 2#100 is set later additionally so the firmware can detect our cycle time)
      NewHandShakeValue := 2#011;

      b_TimeSyncActive := TRUE;

//**********************************************************************************************************************************************************
    CMD_SM_INIT_FINISHED:
      // the safety manager has finished his administration work (e.g. connecting the domains)
      b_ManagerInitialisationFinished := TRUE;

      // optional modules may not be available
      ud_OptionalTimeoutStart := ops.tAbsolute;

      UnsafeScheduler := UnsafeSchedulerSetBusReady;
      us_SetBusReadyState := WaitPDOsSyncron;

//**********************************************************************************************************************************************************
    CMD_SM_FIRST_CONNECT_READY:
      // the safety manager has finished first time connecting the domains
      b_ManagerReadyForSDO := TRUE;

//**********************************************************************************************************************************************************
    CMD_SM_DISCONNECT:
      b_ManagerInitialisationFinished := FALSE;
      b_ManagerReadyForSDO := FALSE;

      // wait again to send bus ready signal
      if ClassState <> _ReinitConfig then
        ClassState := _WaitForSynchronicity;
      end_if;
      UnsafeScheduler := UnsafeSchedulerSetBusReady;
      us_SetBusReadyState := WaitPDOsSyncron;

//**********************************************************************************************************************************************************
    CMD_SM_SDO_TO_MODULE:
#ifdef DO_DEBUG
      DOCheck(pFrame:=(pPara^.aPara[1])$^SDOStdHeader, pCheckStruct:=#SDOWrite);
#endif

      AddSDOToBuffer(p_us_Message := pPara^.aPara[1]$^USINT, us_length := pPara^.aPara[0]$USINT);

//**********************************************************************************************************************************************************
    CMD_SM_TDO_TO_MODULE:
      WriteTDO2Module(pTDO:=(pPara^.aPara[1])$^TDOType);

//**********************************************************************************************************************************************************
    CMD_SM_GET_SAFETY_NUMBER:
      // check if pointer is valid
      if pPara^.aPara[0] then
        ((pPara^.aPara[0])$^UDINT)^ := SafetyNumber;
      end_if;
//**********************************************************************************************************************************************************
    CMD_SM_ADD_INPUT_PDO:
      AddPDOToInputBuffer(ud_p2Buffer         := pPara^.aPara[0]$UDINT
                        , ud_HandleSourceDO   := pPara^.aPara[5]$UDINT
                        , ud_MoveSourceAddr   := pPara^.aPara[1]$UDINT
                        , ud_MoveSourceOffset := pPara^.aPara[6]$UDINT
                        , ud_SafetyNr         := pPara^.aPara[2]$UDINT
                        , b_IsOptional        := pPara^.aPara[4]$BOOL
                        , us_PdoLen           := pPara^.aPara[3]$USINT);

//**********************************************************************************************************************************************************
    CMD_SM_ADD_OUTPUT_PDO:
      // if it's an interface frame, we return the pointer to the second PDO frame which is the interface pdo frame
      if pPara^.aPara[0] = 1 then
        // skip the first PDO
        pResult^.aData[0]$UDINT := GetPointer2PDOBuffer() + MyPDOSize;
        pResult^.aData[4]$UDINT := pPDOReadData$UDINT + MyPDOSize;
        pResult^.aData[8]$UDINT := p_HandlePDORead$UDINT; // Still the same DO Handle
        pResult^.aData[12]$UDINT:= MyPDOSize$UDINT;
        pResult^.aData[8]$UDINT := p_HandlePDORead$UDINT; // Still the same DO Handle
        pResult^.aData[12]$UDINT:= MyPDOSize$UDINT;
      else
        // otherwise just get the pointer to the PDO read data
        pResult^.aData[0]$UDINT := GetPointer2PDOBuffer();
        pResult^.aData[4]$UDINT := pPDOReadData$UDINT;
        pResult^.aData[8]$UDINT := p_HandlePDORead$UDINT;
        pResult^.aData[12]$UDINT:= 0$UDINT;
        pResult^.aData[8]$UDINT := p_HandlePDORead$UDINT;
        pResult^.aData[12]$UDINT:= 0$UDINT;
      end_if;

      // p_HandlePDORead

      pResult^.uiLng := 16;

//**********************************************************************************************************************************************************
    CMD_SM_REMOVE_INPUT_PDO:
      // we lost connection to other systems => we have to initialize again! remove old input PDOs

      if ui_cnt_PDOInputBuffer then
        // save the old state of the class and set it temporarily to "module not found" to prevent update rt from crashing
        OldClassState := ClassState;
        ClassState := _ModuleNotFound;

        // search for the PDO
        Found := FALSE;
        pPDOInputBuffer := #aPDOInputBuffer[0];
        for i := 0 to (ui_cnt_PDOInputBuffer-1) do
          if pPDOInputBuffer^.ud_p2Buffer = pPara^.aPara[0]$UDINT then
            Found := TRUE;
            exit;
          end_if;

          pPDOInputBuffer += sizeof(PDOInputBuffer);
        end_for;

        // if we found the PDO => remove it from memory (move the memory behind the found PDO over the place of the found PDO)
        if Found then
          // if it's last entry (no entries have to be moved) => we only have to copy some memory if it's not the last
          if i < (ui_cnt_PDOInputBuffer-1) then
            for j := i to (ui_cnt_PDOInputBuffer-2) do
              aPDOInputBuffer[j] := aPDOInputBuffer[j+1];
            end_for;
          end_if;
          ui_cnt_PDOInputBuffer -= 1;
        else
          LogError("@ZZZZ (SafetyCDIAS_Base::State::NewInst) CMD_SM_REMOVE_INPUT_PDO failed! Couldn't find specified PDO!");
        end_if;

        // restore old class state
        ClassState := OldClassState;
      else
        LogError("@ZZZZ (SafetyCDIAS_Base::State::NewInst) CMD_SM_REMOVE_INPUT_PDO failed! No input PDOs found!");
      end_if;

//*****************************************************************************
//** COMMANDS FROM OTHER SAFETYMODULES                                       **
//*****************************************************************************

//**********************************************************************************************************************************************************
    CMD_SM_ADD_SDO_TO_BUFFER:
      sd_retval := AddSDOToBuffer(p_us_message:=pPara^.aPara[0]$^USINT, us_length:=pPara^.aPara[1]$USINT);
      if sd_retval then
        ret_code := 1$IprStates; //means iprStates::ERROR but a server error also exists
      end_if;

      pResult^.aData[0]$DINT := sd_retval;

//**********************************************************************************************************************************************************
    CMD_SM_WRITE_TDO_TO_MODULE:
      WriteTDO2Module(pTDO:=pPara^.aPara[0]$^TDOType);

//**********************************************************************************************************************************************************
    CMD_SM_CONFIG_SAFETY_CPU:
      pResult^.aData[0]$UDINT := ConfigSafetyCpu();

//**********************************************************************************************************************************************************
    CMD_SM_CONFIG_SAFETY_INPUT:
      pResult^.aData[0]$UDINT := ConfigSafetyInput(ud_SafeNrCPU         := pPara^.aPara[0]$HDINT
                                                 , ud_thisp             := pPara^.aPara[1]$UDINT
                                                 , p_PDOBuffer          := pPara^.aPara[2]$^UDINT
                                                 , pMoveActive          := pPara^.aPara[3]$^PDOMoveState
                                                 , p_ud_HandleSourceDO  := pPara^.aPara[5]$^UDINT
                                                 , p_ud_MoveSourceAddr  := pPara^.aPara[4]$^UDINT
                                                 , p_ud_MoveSourceOffset:= pPara^.aPara[6]$^UDINT
                                                 );

//**********************************************************************************************************************************************************
    CMD_SM_CONFIG_SAFETY_OUTPUT:
      pResult^.aData[0]$UDINT := ConfigSafetyOutput(ud_SafeNrCPU        := pPara^.aPara[0]$HDINT
                                                  , ud_thisp            := pPara^.aPara[1]$UDINT
                                                  , ud_p_PDOBuffer      := pPara^.aPara[2]$UDINT
                                                  , pObject             := pPara^.aPara[3]$^PathInfoType
                                                  , pMoveActive         := pPara^.aPara[4]$^PDOMoveState
                                                  , ud_HandleSourceDO   := pPara^.aPara[7]$UDINT
                                                  , ud_MoveSourceAddr   := pPara^.aPara[5]$UDINT
                                                  , ud_MoveSourceOffset := pPara^.aPara[8]$UDINT
                                                  , b_IsOptional        := pPara^.aPara[6]$BOOL
                                                  );

//**********************************************************************************************************************************************************
    CMD_SM_REMOVE_CPU_FROM_TABLE:
      RemoveCPUFromTable(ud_SafetyNr := pPara^.aPara[0]$HDINT);

//**********************************************************************************************************************************************************
    CMD_SM_GET_MODULE_TYPE:
      pResult^.aData[0]$UDINT := SM_TYPE_SAFETY_MODULE;

//**********************************************************************************************************************************************************
    CMD_SM_DEACTIVATE_MOVE_CMD:
      // check if it's for input (1) or output (0)
      if pPara^.aPara[0] then
        b_MoveCommandInputActive  := _Inactive;
      else
        b_MoveCommandOutputActive := _Inactive;
      end_if;

//**********************************************************************************************************************************************************
    CMD_SM_MODULE_REINIT:
      if b_ReInitMarker then
        if GetModuleID() = CSCP01x_ID then

          // delete request
          LastRequest := _NoOpenRequest;
          ud_AsyComRetryCounter := 0; // reset retry counter

          // remove the cpu from all classes, which use it
          ResetConfig();

          if UnsafeScheduler <> UnsafeSchedulerSetBusReady then
            us_SetBusReadyState := WaitPDOsSyncron;
            UnsafeScheduler := UnsafeSchedulerSetBusReady;
          end_if;

          MaxVarsPerReadPackage   := 0;
          ReadFramesNeeded        := 0;
          MaxVarsPerWritePackage  := 0;
          WriteFramesNeeded       := 0;

          ClassState := _ReinitConfig;
          b_GetNewConfiguration := TRUE;
        end_if;

        b_ReInitMarker := FALSE;
      end_if;

//**********************************************************************************************************************************************************
    CMD_SM_POST_INIT_FINISHED:

      b_PostInitPassed := TRUE;

      if ( State.uiIO_Flags = 0 ) then

        // get configuration if module is configured

        // get state via SDO communication
        sd_retval := SDOStdRequ ( us_Command      := SDO_COMMAND_GET_STATE
                                , p_us_RespData   := ( #GetStateResp )$^USINT
                                , us_RespLength   := sizeof(GetStateResponseType)
                                );

        // the cpu is configured, load the new configuration
        if ( sd_retval = 0 ) &
           (GetStateResp.ConfigState <> CFG_STATE_UNKNOWN) &
           (GetStateResp.ConfigState <> CFG_STATE_INVALID) &
           (GetStateResp.ConfigState <> CFG_STATE_NOT_CONFIGURED) then

          //get configuration from safe CPU and build routing tables
          GetRoutingData();
        else
          //get configuration from safe CPU and build routing tables later in background
          b_GetNewConfiguration := FALSE;

            // next time we check for the configured state of the cpu
          b_CheckConfigured     := TRUE;

          // check again in background
          ClassState            := _ReinitConfig;
        end_if;
      end_if;

//**********************************************************************************************************************************************************
  CMD_GET_HARDWARE_DIAGNOSIS:
    //Set Errors

    ret_code := 1$IprStates; //means iprStates::ERROR but a server error also exists

    pResult^.aData[0]$t_HWCGetHardwareDiagnosisOut.retcode           := _HWC_RETVAL_ERROR_CLASS_NOT_ONLINE;

    //Return State and Device ID and Kennung of placed module --------------------------------
    if State.uiIO_Flags.WrongHW = 1 then
      pResult^.aData$t_HWCGetHardwareDiagnosisOut.ClassState := _WrongHardware;
      pResult^.aData[0]$t_HWCGetHardwareDiagnosisOut.retcode := _HWC_RETVAL_ERROR_WRONG_HARDWARE;
    elsif State.uiIO_Flags.NoHW = 1 then
      pResult^.aData$t_HWCGetHardwareDiagnosisOut.ClassState := _NoHardware;
      pResult^.aData[0]$t_HWCGetHardwareDiagnosisOut.retcode := _HWC_RETVAL_ERROR_NO_HARDWARE;
    elsif State.uiIO_Flags.NoCalibration = 1 then
      pResult^.aData$t_HWCGetHardwareDiagnosisOut.ClassState := _NoCalibDataFound;
      pResult^.aData[0]$t_HWCGetHardwareDiagnosisOut.retcode := _HWC_RETVAL_ERROR_NO_CALIB_DATA_FOUND;
    end_if;

    pResult^.aData$t_HWCGetHardwareDiagnosisOut.ud_DeviceID := GetModuleID();
    pResult^.aData$t_HWCGetHardwareDiagnosisOut.ud_Variante := GetKennung();

    //-----------------------------------------------------------------------------------------

    // Only respond if the class is online
    if State.uiIO_Flags = 0 then
      pResult^.aData$t_HWCGetHardwareDiagnosisOut.ClassState := _ClassOk;
      ptmpStr := pPara^.aPara[0]$t_HWCGetHardwareDiagnosisIn.pStr_HardewareTreeEntry;

      // Check if position pointers strings are valid
      if ptmpStr & p_ObjectPath then

        // Length is 2 byte for ptmpStr and 1 byte for p_ObjectPath
        if (ptmpStr)$^UINT^ > 0 & (ptmpStr)$^UINT^ = (p_ObjectPath)$^USINT^ then // Check if length if positionstring is valid and equal

          if _memcmp(ptr1:=ptmpStr+2, ptr2:=p_ObjectPath+1, cntr:= (ptmpStr)$^UINT^) = 0 then  // Compare strings , 2 bytes length for ptmpStr, 1 byte length for p_ObjectPath

            ret_code := READY;
            pResult^.aData[0]$t_HWCGetHardwareDiagnosisOut.retcode           := _HWC_RETVAL_OK;
            pResult^.aData[0]$t_HWCGetHardwareDiagnosisOut.pStr_DeviceName   := NIL;
            pResult^.aData[0]$t_HWCGetHardwareDiagnosisOut.pStr_VendorName   := NIL;
            pResult^.aData[0]$t_HWCGetHardwareDiagnosisOut.ud_VendorID       := 0;

            // Get Serialno -----------------------------------------------------------------------------------------
            ud_StrSize := SerialNoStr.GetLength() ;
            pResult^.aData[0]$t_HWCGetHardwareDiagnosisOut.pStr_SerialNo     := NIL;

            if ud_StrSize then

              if (ud_StrSize < sizeof(a_SerialNo)) then // < to account for 0 termination
                // Copy complete string
                SerialNoStr.GetDataAt(pData:=#a_SerialNo[0], udSize:=ud_StrSize, udAt:=0);
                a_SerialNo[ud_StrSize] := 0; // 0 termination
              else
                // Copy part string
                SerialNoStr.GetDataAt(pData:=#a_SerialNo[0], udSize:=sizeof(a_SerialNo)-1, udAt:=0);
                a_SerialNo[sizeof(a_SerialNo)-1] := 0; // 0 termination
              end_if;
              pResult^.aData[0]$t_HWCGetHardwareDiagnosisOut.pStr_SerialNo     := #a_SerialNo[0];
            end_if;
            // ----------------------------------------------------------------------------------------------------------

            pResult^.aData[0]$t_HWCGetHardwareDiagnosisOut.pStr_OrderingNo   := NIL;
            pResult^.aData[0]$t_HWCGetHardwareDiagnosisOut.ud_LicenseNo      := 0;

            // Get Hardwareversion --------------------------------------------------------------------------------------
            pResult^.aData[0]$t_HWCGetHardwareDiagnosisOut.hd_HWVersion := 0;
            if MasterConnect.I2CReadOneByte(AdressCDIAS:=(Place*16#100)$UINT+CDIAS_EEPROM_OFFSET_HWVERSION, pData:=#us_temp) = 0 then
              pResult^.aData[0]$t_HWCGetHardwareDiagnosisOut.hd_HWVersion := us_temp;
            end_if;

            // Get Variante --------------------------------------------------------------------------------------
              pResult^.aData[0]$t_HWCGetHardwareDiagnosisOut.ud_Variante := 0;
            if MasterConnect.I2CReadOneByte(AdressCDIAS:=(Place*16#100)$UINT+CDIAS_EEPROM_OFFSET_VARIANTE, pData:=#us_temp) = 0 then
              pResult^.aData[0]$t_HWCGetHardwareDiagnosisOut.ud_Variante := us_temp;
            end_if;

            // Get FPGA Version -----------------------------------------------------------------------------------------
            pResult^.aData[0]$t_HWCGetHardwareDiagnosisOut.hd_FPGAVersion := FPGA_Version;

            //Get Safetynumber ------------------------------------------------------------------------------------------
            pResult^.aData[0]$t_HWCGetHardwareDiagnosisOut.hd_SafetyNumber := SafetyNumber;

            //Get FW Version --------------------------------------------------------------------------------------------
            GetFWVersion(pData:=#a_FWVersion[0],sizeof(a_FWVersion));
            pResult^.aData$t_HWCGetHardwareDiagnosisOut.pStr_FWVersion := #a_FWVersion[0];

            // -----------------------------------------------------------------------------------------------------------

            pResult^.aData[0]$t_HWCGetHardwareDiagnosisOut.ud_Place          := Place;
            pResult^.aData[0]$t_HWCGetHardwareDiagnosisOut.ud_reserved_size  := 0;
            pResult^.aData[0]$t_HWCGetHardwareDiagnosisOut.pud_reserved      := NIL;
            pResult^.aData[0]$t_HWCGetHardwareDiagnosisOut.ud_user_size      := 0;
            pResult^.aData[0]$t_HWCGetHardwareDiagnosisOut.pud_user          := NIL;
            pResult^.aData[0]$t_HWCGetHardwareDiagnosisOut.p_DynExtList      := NIL;
          end_if;

        end_if;

      end_if;
//      else
//        pResult^.aData[0]$t_HWCGetHardwareDiagnosisOut.retcode           := _HWC_RETVAL_ERROR_CLASS_NOT_ONLINE;
    end_if;

//**********************************************************************************************************************************************************
  else
    // needed for required handling
    ret_code := HwBaseCDIAS::NewInst(pPara, pResult);
//**********************************************************************************************************************************************************
  END_CASE;

END_FUNCTION

FUNCTION VIRTUAL SafetyCDIAS_Base::ShowProjectRevision
// to overload in cscp class
END_FUNCTION

FUNCTION SafetyCDIAS_Base::DOCheck
	VAR_INPUT
		pFrame 	      : ^SDOStdHeader;
		pCheckStruct 	: ^t_DataObjectCheck;
	END_VAR
  VAR
  	DOCheckHeader : SDOStdHeader;
    ActTime       : UDINT;
  END_VAR

  // check if input parameters are correct
  if pFrame & pFrame^.Len & pCheckStruct then
    DOCheckHeader := pFrame^;

    // only if we got a different frame
    if DOCheckHeader <> pCheckStruct^.LastHeader then
      ActTime := OS_READMICROSEC();

      pCheckStruct^.TimeDiff := ActTime - pCheckStruct^.LastTime;

      if pCheckStruct^.TimeDiff > pCheckStruct^.TimeDiffMax then
        if pCheckStruct^.TimeDiffMax = 0 then
          pCheckStruct^.TimeDiffMax := 1;
        else
          pCheckStruct^.TimeDiffMax := pCheckStruct^.TimeDiff;
        end_if;
      end_if;

      if pCheckStruct^.TimeDiff < pCheckStruct^.TimeDiffMin then
        pCheckStruct^.TimeDiffMin := pCheckStruct^.TimeDiff;
      end_if;

      pCheckStruct^.LastTime := ActTime;
    else
      // if it's the same frame again: problem!
      pCheckStruct^.SameFrameCnt += 1;
    end_if;
    pCheckStruct^.LastHeader := DOCheckHeader;
  end_if;

END_FUNCTION

FUNCTION VIRTUAL SafetyCDIAS_Base::CalcPDOLength
	VAR_INPUT
		BoolVarNo 	: UDINT;
		DintVarNo 	: UDINT;
	END_VAR
	VAR_OUTPUT
		PdoLen 	    : USINT;
	END_VAR
  VAR
    PayLoad     : USINT;
  END_VAR

  // we have at least the header
  PdoLen  := sizeof(PDOType) - sizeof(PDOType.DataAndCopy);
  PayLoad := 0;

  // now add some space for the needed data
  if BoolVarNo then
    // 1 byte (type + number of values) + 1 byte index + 2 bits for every value (4 per byte)
    PayLoad += 2 + ((BoolVarNo$USINT + 3) / 4);

    // make the it 2 byte aligned (if it isn't already) => only if no dint variables, otherwise it is done one at the DINT variables
    if (PayLoad MOD 2) & (DintVarNo = 0) then
      PayLoad := PayLoad + (2 - (PayLoad MOD 2)); //increase memory, up to a value, which could be divided by 2
    end_if;
  end_if;

  if DintVarNo then
    // 1 byte (type + number of values) + 1 byte index + 1 byte errorflags per 8 values + 4 byte for every value
    PayLoad += 2 + (((DintVarNo$USINT - 1 ) / 8) + 1) + DintVarNo$USINT * 4;

    // make the it 2 byte aligned (if it isn't already)
    if (PayLoad MOD 2) then
      PayLoad := PayLoad + (2 - (PayLoad MOD 2)); //increase memory, up to a value, which could be divided by 2
    end_if;
  end_if;

  // duplicate it
  PayLoad *= 2;

  // add it to the total length
  PdoLen += PayLoad;

END_FUNCTION

FUNCTION VIRTUAL SafetyCDIAS_Base::AddModuleToCfg
	VAR_INPUT
		ModuleCfg : t_ModuleCfg;
	END_VAR
	VAR_OUTPUT
		retcode 	: DINT;
	END_VAR
  VAR
    pHelp     : ^t_ModuleListElem;
  END_VAR

  retcode := 0;

  if pFirstModuleCfg = NIL then
    pFirstModuleCfg$pVoid := To_StdLib.Malloc(size:=sizeof(t_ModuleListElem));
    pHelp := pFirstModuleCfg;
  else
    pHelp := pFirstModuleCfg;
    // if searched path has been found, we already got this module in our list
    if (ModuleCfg.PathLen = pHelp^.ModuleInfo.PathLen) & (To_StdLib.MemCmp(dest:= ModuleCfg.pPath, source:= pHelp^.ModuleInfo.pPath , size:= ModuleCfg.PathLen) = 0) then
      // already in buffer => leave function
      return;
    end_if;
    while pHelp^.pNext <> NIL do
      // if searched path has been found, we already got this module in our list
      if (ModuleCfg.PathLen = pHelp^.ModuleInfo.PathLen) & (To_StdLib.MemCmp(dest:= ModuleCfg.pPath, source:= pHelp^.ModuleInfo.pPath , size:= ModuleCfg.PathLen) = 0) then
        // already in buffer => leave function
        return;
      else
        pHelp := pHelp^.pNext;
      end_if;
    end_while;

    // if searched path has been found, we already got this module in our list
    if (ModuleCfg.PathLen = pHelp^.ModuleInfo.PathLen) & (To_StdLib.MemCmp(dest:= ModuleCfg.pPath, source:= pHelp^.ModuleInfo.pPath , size:= ModuleCfg.PathLen) = 0) then
      // already in buffer => leave function
      return;
    else
      pHelp^.pNext$pvoid := To_StdLib.Malloc(size:=sizeof(t_ModuleListElem));
      pHelp := pHelp^.pNext;
    end_if;
  end_if;

  if pHelp <> NIL then
    // allocate memory for the module path
    pHelp^.ModuleInfo.pPath$pVoid := To_StdLib.Malloc(size:=ModuleCfg.PathLen);
    if pHelp^.ModuleInfo.pPath = NIL then
      ClassState := _MemAllocFailed;
      retcode := -1;
      return;
    end_if;

    _memcpy(ptr1:=pHelp^.ModuleInfo.pPath, ptr2:=ModuleCfg.pPath, cntr:=ModuleCfg.PathLen);

    // allocate memory for the module path
    pHelp^.ModuleInfo.pCompPath$pVoid := To_StdLib.Malloc(size:=ModuleCfg.CompPathLen);
    if pHelp^.ModuleInfo.pCompPath = NIL then
      ClassState := _MemAllocFailed;

      retcode := -1;
      return;
    end_if;

    _memcpy(ptr1:=pHelp^.ModuleInfo.pCompPath, ptr2:=ModuleCfg.pCompPath, cntr:=ModuleCfg.CompPathLen);

    pHelp^.ModuleInfo.Info        := ModuleCfg.Info;
    pHelp^.ModuleInfo.SafetyNbr   := ModuleCfg.SafetyNbr;
    pHelp^.ModuleInfo.InterfaceCRC:= ModuleCfg.InterfaceCRC;
    pHelp^.ModuleInfo.DestCRCNo   := ModuleCfg.DestCRCNo;
    phelp^.ModuleInfo.pDestCRCs   := ModuleCfg.pDestCRCs;
    pHelp^.ModuleInfo.PathLen     := ModuleCfg.PathLen;
    pHelp^.ModuleInfo.CompPathLen := ModuleCfg.CompPathLen;
    pHelp^.ModuleInfo.PdoOutLen   := ModuleCfg.PdoOutLen;

    pHelp^.pNext                  := NIL;

    ModuleCfgNo += 1;
  else
    ClassState := _MemAllocFailed;
    retcode := -1;
    return;
  end_if;

END_FUNCTION

FUNCTION VIRTUAL SafetyCDIAS_Base::AddPdoToCfg
	VAR_INPUT
		PdoCfg 	: t_PdoCfg;
	END_VAR
	VAR_OUTPUT
		retcode 	: DINT;
	END_VAR
  VAR
    pHelp : ^t_PdoListElem;
  END_VAR

  retcode := 0;

  if pFirstPdoCfg = NIL then
    pFirstPdoCfg$pVoid := To_StdLib.Malloc(size:=sizeof(t_PdoListElem));
    pHelp := pFirstPdoCfg;
  else
    pHelp := pFirstPdoCfg;
    // if searched path has been found, we already got this pdo in our list
    if (PdoCfg.SourcePathLen = pHelp^.PdoInfo.SourcePathLen) & (PdoCfg.DestPathLen = pHelp^.PdoInfo.DestPathLen) &
      (PdoCfg.InterfaceCRC = pHelp^.PdoInfo.InterfaceCRC) &
      (To_StdLib.MemCmp(dest:= PdoCfg.pSourcePath, source:= pHelp^.PdoInfo.pSourcePath , size:= PdoCfg.SourcePathLen) = 0) &
      (To_StdLib.MemCmp(dest:= PdoCfg.pDestPath,   source:= pHelp^.PdoInfo.pDestPath   , size:= PdoCfg.DestPathLen  ) = 0) then
      // already in buffer => leave function
      return;
    end_if;
    while pHelp^.pNext <> NIL do
      // if searched path has been found, we already got this pdo in our list
      if (PdoCfg.SourcePathLen = pHelp^.PdoInfo.SourcePathLen) & (PdoCfg.DestPathLen = pHelp^.PdoInfo.DestPathLen) &
        (PdoCfg.InterfaceCRC = pHelp^.PdoInfo.InterfaceCRC) &
        (To_StdLib.MemCmp(dest:= PdoCfg.pSourcePath, source:= pHelp^.PdoInfo.pSourcePath , size:= PdoCfg.SourcePathLen) = 0) &
        (To_StdLib.MemCmp(dest:= PdoCfg.pDestPath,   source:= pHelp^.PdoInfo.pDestPath   , size:= PdoCfg.DestPathLen  ) = 0) then
        // already in buffer => leave function
        return;
      else
        pHelp := pHelp^.pNext;
      end_if;
    end_while;

    // if searched path has been found, we already got this pdo in our list
    if (PdoCfg.SourcePathLen = pHelp^.PdoInfo.SourcePathLen) & (PdoCfg.DestPathLen = pHelp^.PdoInfo.DestPathLen) &
      (PdoCfg.InterfaceCRC = pHelp^.PdoInfo.InterfaceCRC) &
      (To_StdLib.MemCmp(dest:= PdoCfg.pSourcePath, source:= pHelp^.PdoInfo.pSourcePath , size:= PdoCfg.SourcePathLen) = 0) &
      (To_StdLib.MemCmp(dest:= PdoCfg.pDestPath,   source:= pHelp^.PdoInfo.pDestPath   , size:= PdoCfg.DestPathLen  ) = 0) then
      // already in buffer => leave function
      return;
    else
      pHelp^.pNext$pvoid := To_StdLib.Malloc(size:=sizeof(t_PdoListElem));
      pHelp := pHelp^.pNext;
    end_if;
  end_if;

  if pHelp <> NIL then
    // allocate memory for the module source path
    pHelp^.PdoInfo.pSourcePath$pVoid := To_StdLib.Malloc(size:=PdoCfg.SourcePathLen);
    if pHelp^.PdoInfo.pSourcePath = NIL then
      ClassState := _MemAllocFailed;
      retcode := -1;
      return;
    end_if;

    _memcpy(ptr1:=pHelp^.PdoInfo.pSourcePath, ptr2:=PdoCfg.pSourcePath, cntr:=PdoCfg.SourcePathLen);

    // allocate memory for the module source path
    pHelp^.PdoInfo.pDestPath$pVoid := To_StdLib.Malloc(size:=PdoCfg.DestPathLen);
    if pHelp^.PdoInfo.pDestPath = NIL then
      ClassState := _MemAllocFailed;
      retcode := -1;
      return;
    end_if;

    _memcpy(ptr1:=pHelp^.PdoInfo.pDestPath, ptr2:=PdoCfg.pDestPath, cntr:=PdoCfg.DestPathLen);

    pHelp^.PdoInfo.Info           := PdoCfg.Info;
    pHelp^.PdoInfo.InterfaceCRC   := PdoCfg.InterfaceCRC;
    pHelp^.PdoInfo.SourcePathLen  := PdoCfg.SourcePathLen;
    pHelp^.PdoInfo.DestPathLen    := PdoCfg.DestPathLen;
    // length is only zero for non-interface pdos
    if PdoCfg.Info.IsInterfacePDO = FALSE then
      pHelp^.PdoInfo.PdoLen       := 0;   // the length is determined later in method CreateAndSendCfg
    else
      pHelp^.PdoInfo.PdoLen       := PdoCfg.PdoLen;
    end_if;
    pHelp^.PdoInfo.PDO_ID         := 255; // the ID is assigned later by the safety manager of the master domain
    pHelp^.pNext                  := NIL;

    PdoCfgNo += 1;
  else
    ClassState  := _MemAllocFailed;
    retcode     := -1;
    return;
  end_if;

END_FUNCTION

FUNCTION VIRTUAL SafetyCDIAS_Base::AddSlaveToCfg
	VAR_INPUT
		pModule 	    : ^PathInfoType;
		b_IsOptional 	: BOOL;
		b_IsInterface : BOOL;
		InterfaceCRC 	: HDINT;
	END_VAR
  VAR
    pHelp         : ^t_SlaveListElem;
  END_VAR

  if pFirstSlaveCfg = NIL then
    pFirstSlaveCfg$pVoid := To_StdLib.Malloc(size:=sizeof(t_SlaveListElem));
    pHelp := pFirstSlaveCfg;
  else
    pHelp := pFirstSlaveCfg;
    while pHelp^.pNext <> NIL do
      //if searched path is found, we already got this module in our list
      if (pModule^.ui_PathCompLen = pHelp^.SlaveInfo.CompPathLen) &
        (To_StdLib.MemCmp(dest:= pModule^.p_us_PathComp, source:= pHelp^.SlaveInfo.pCompPath , size:= pModule^.ui_PathCompLen) = 0) then
        // already in buffer => leave function
        return;
      else
        pHelp := pHelp^.pNext;
      end_if;
    end_while;

    //if searched path is found, we already got this module in our list
    if (pModule^.ui_PathCompLen = pHelp^.SlaveInfo.CompPathLen) &
      (To_StdLib.MemCmp(dest:= pModule^.p_us_PathComp, source:= pHelp^.SlaveInfo.pCompPath , size:= pModule^.ui_PathCompLen) = 0) then
      // already in buffer => leave function
      return;
    end_if;

    pHelp^.pNext$pvoid := To_StdLib.Malloc(size:=sizeof(t_SlaveListElem));
    pHelp := pHelp^.pNext;
  end_if;

  if pHelp <> NIL then
    // allocate memory for the module path
    pHelp^.SlaveInfo.PathLen := pModule^.p_us_Path^$UINT + 2;
    pHelp^.SlaveInfo.pPath$pVoid := To_StdLib.Malloc(size:=pHelp^.SlaveInfo.PathLen);
    if pHelp^.SlaveInfo.pPath = NIL then
      ClassState := _MemAllocFailed;
      LogError("@ZZZZ (SafetyCDIAS_Base::AddSlaveToCfg) Error: Failed to allocate memory for the module path");
      return;
    end_if;

    _memcpy(ptr1:=pHelp^.SlaveInfo.pPath, ptr2:=pModule^.p_us_Path, cntr:=pHelp^.SlaveInfo.PathLen);

    // allocate memory for the module path
    pHelp^.SlaveInfo.CompPathLen := pModule^.ui_PathCompLen;
    pHelp^.SlaveInfo.pCompPath$pVoid := To_StdLib.Malloc(size:=pHelp^.SlaveInfo.CompPathLen);
    if pHelp^.SlaveInfo.pCompPath = NIL then
      ClassState := _MemAllocFailed;
      LogError("@ZZZZ (SafetyCDIAS_Base::AddSlaveToCfg) Error: Failed to allocate memory for the compressed module path");
      return;
    end_if;

    _memcpy(ptr1:=pHelp^.SlaveInfo.pCompPath, ptr2:=pModule^.p_us_PathComp, cntr:=pHelp^.SlaveInfo.CompPathLen);

    pHelp^.SlaveInfo.Info             := 0;
    pHelp^.SlaveInfo.Info.IsOptional  := b_IsOptional;
    pHelp^.SlaveInfo.Info.IsInterface := b_IsInterface;

    pHelp^.SlaveInfo.InterfaceCRC     := InterfaceCRC;

    pHelp^.pNext                      := NIL;

    SlaveCfgNo += 1;
  else
    ClassState := _MemAllocFailed;
    LogError("@ZZZZ (SafetyCDIAS_Base::AddSlaveToCfg) Error: Failed to allocate memory for the new list-element");
    return;
  end_if;

END_FUNCTION

FUNCTION VIRTUAL SafetyCDIAS_Base::FreeCfgLists
  VAR
    pHelpModule : ^t_ModuleListElem;
    pHelpPdo    : ^t_PdoListElem;
    pHelpSlave  : ^t_SlaveListElem;
//    pHelpUnsafeVar : ^t_UnsafeVarListElem;
  END_VAR

  // while we got module cfgs
  while pFirstModuleCfg do
    pHelpModule := pFirstModuleCfg;
    pFirstModuleCfg := pFirstModuleCfg^.pNext;

    if pHelpModule^.ModuleInfo.pDestCRCs then
      To_StdLib.Free(pHelpModule^.ModuleInfo.pDestCRCs);
    end_if;
    To_StdLib.Free(pHelpModule^.ModuleInfo.pPath);
    To_StdLib.Free(pHelpModule^.ModuleInfo.pCompPath);
    To_StdLib.Free(pHelpModule);
  end_while;
  pFirstModuleCfg := NIL;
  ModuleCfgNo     := 0;

  // while we got pdo cfgs
  while pFirstPdoCfg do
    pHelpPdo := pFirstPdoCfg;
    pFirstPdoCfg := pFirstPdoCfg^.pNext;

    To_StdLib.Free(pHelpPdo^.PdoInfo.pSourcePath);
    To_StdLib.Free(pHelpPdo^.PdoInfo.pDestPath);
    To_StdLib.Free(pHelpPdo);
  end_while;
  pFirstPdoCfg := NIL;
  PdoCfgNo := 0;

  // while we got slave cfgs
  while pFirstSlaveCfg do
    pHelpSlave := pFirstSlaveCfg;
    pFirstSlaveCfg := pFirstSlaveCfg^.pNext;

    To_StdLib.Free(pHelpSlave^.SlaveInfo.pPath);
    To_StdLib.Free(pHelpSlave^.SlaveInfo.pCompPath);
    To_StdLib.Free(pHelpSlave);
  end_while;
  pFirstSlaveCfg := NIL;
  SlaveCfgNo := 0;

// memory is freed by safety manager
//  // while we got unsafevar cfgs
//  while pFirstUnsafeCfg do
//    pHelpUnsafeVar := pFirstUnsafeCfg;
//    pFirstUnsafeCfg := pFirstUnsafeCfg^.pNext;
//
//    To_StdLib.Free(pHelpUnsafeVar^.UnsafeVarInfo.pName);
//    To_StdLib.Free(pHelpUnsafeVar);
//  end_while;
//  pFirstUnsafeCfg := NIL;
//  UnsafeCfgNo := 0;

  // reduze size of config mem used to 4 (only safety number of cpu module)
  ConfigMemSizeUsed := 4;

END_FUNCTION

FUNCTION VIRTUAL SafetyCDIAS_Base::CreateAndSendCfg
  VAR
    pHelpModule   : ^t_ModuleListElem;
    pHelpPdo      : ^t_PdoListElem;
    pHelpSlave    : ^t_SlaveListElem;
    pCfg          : ^void;
    TmpPathLen    : UINT;
		MyPara 	      : CmdStruct;
		MyResult	    : results;
    AddConfigSize : UDINT;
  END_VAR

(*
    Memory structure:
      4 Byte: SafetyNumber of CPU (is already there from initialisation in CSCP011_IM::InitSafeModule)
      1 Byte: Number of module configurations which are following
      for every module configuration (first is always the CPU itself)
        1 Byte: Info
        4 Byte: Interface Frame Source SafetyNumber (0 if it is no source for interface frames)
        4 Byte: Interface Frame CRC
        1 Byte: Number of destination inferface frame CRCs
        x Byte: Destination interface frame CRCs (number * sizeof(HDINT)
        2 Byte: Length of hardware path
        x Byte (depending on length in the 2 byte before): Hardwarepath
        2 Byte: Length of compressed hardware path
        x Byte (depending on length in the 2 byte before): Compressed Hardwarepath
        1 Byte: PDO out length for this module
      1 Byte: Number of pdo configurations which are following
      for every PDO configuration
        1 Byte: PDO length
        1 Byte: Interface frame info
        4 Byte: Interface CRC
        2 Byte: Length of source hardware path
        x Byte (depending on length in the 2 byte before): Hardwarepath of source
        2 Byte: Length of destination hardware path
        x Byte (depending on length in the 2 byte before): Hardwarepath of destination
      1 Byte: Number of slave configurations which are following
      for every slave configuration
        1 Byte: Info
        4 Byte: InterfaceCRC
        2 Byte: Length of hardware path
        x Byte (depending on length in the 2 byte before): Hardwarepath
        2 Byte: Length of compressed hardware path
        x Byte (depending on length in the 2 byte before): Compressed Hardwarepath
*)

  // check if there is memory and if the only thing inside is the safety number
  if pConfigMem & (ConfigMemSizeUsed = 4) then
    // pCfg points to the next memory we have to write to => set it to the memory after the safety number
    pCfg := pConfigMem + ConfigMemSizeUsed;

    // add all module configurations to memory
    if pFirstModuleCfg then
      // add number of module configurations to memory (no need to check the memory here, because already 512 bytes are allocated)
      pCfg^$USINT       := ModuleCfgNo;
      pCfg              += sizeof(USINT);
      ConfigMemSizeUsed += sizeof(USINT);

      pHelpModule := pFirstModuleCfg;
      // go through list
      while pHelpModule do
        // add the elements

        // check if we have enough memory to add the next module
        AddConfigSize := sizeof(BSINT) + sizeof(HDINT) + sizeof(HDINT) + sizeof(UINT) + pHelpModule^.ModuleInfo.PathLen + sizeof(UINT) + pHelpModule^.ModuleInfo.CompPathLen + sizeof(USINT);
        if pHelpModule^.ModuleInfo.Info.IsInterfaceDest then
          AddConfigSize += sizeof(USINT) + pHelpModule^.ModuleInfo.DestCRCNo * sizeof(HDINT);
        end_if;

        pCfg := CheckConfigMemSize(AddConfigSize);
        if pCfg = NIL then
          // error message already logged by function
          return;
        end_if;

        // info
        pCfg^$BSINT := pHelpModule^.ModuleInfo.Info;
        pCfg              += sizeof(BSINT);
        ConfigMemSizeUsed += sizeof(BSINT);

        // safety number of interface frame source (if it is one)
        pCfg^$HDINT := pHelpModule^.ModuleInfo.SafetyNbr;
        pCfg              += sizeof(HDINT);
        ConfigMemSizeUsed += sizeof(HDINT);

        // interface CRC of interface frame
        pCfg^$HDINT := pHelpModule^.ModuleInfo.InterfaceCRC;
        pCfg              += sizeof(HDINT);
        ConfigMemSizeUsed += sizeof(HDINT);

        // if its also interface frame destination send the corresponding interface CRCs
        if pHelpModule^.ModuleInfo.Info.IsInterfaceDest then
          TmpPathLen := pHelpModule^.ModuleInfo.DestCRCNo; // save some time with this local variable
          pCfg^$USINT := TmpPathLen$USINT;
          pCfg              += sizeof(USINT);
          ConfigMemSizeUsed += sizeof(USINT);

          _memcpy(ptr1:=pCfg, ptr2:=pHelpModule^.ModuleInfo.pDestCRCs, cntr:=TmpPathLen * sizeof(HDINT));
          pCfg += TmpPathLen * sizeof(HDINT);
          ConfigMemSizeUsed += TmpPathLen * sizeof(HDINT);
        end_if;

        // uncompressed module path
        TmpPathLen := pHelpModule^.ModuleInfo.PathLen; // save some time with this local variable
        pCfg^$UINT := TmpPathLen;
        pCfg              += sizeof(UINT);
        ConfigMemSizeUsed += sizeof(UINT);

        _memcpy(ptr1:=pCfg, ptr2:=pHelpModule^.ModuleInfo.pPath, cntr:=TmpPathLen);
        pCfg += TmpPathLen;
        ConfigMemSizeUsed += TmpPathLen;

        // compressed module path
        TmpPathLen := pHelpModule^.ModuleInfo.CompPathLen; // save some time with this local variable
        pCfg^$UINT := TmpPathLen;
        pCfg              += sizeof(UINT);
        ConfigMemSizeUsed += sizeof(UINT);

        _memcpy(ptr1:=pCfg, ptr2:=pHelpModule^.ModuleInfo.pCompPath, cntr:=TmpPathLen);
        pCfg += TmpPathLen;
        ConfigMemSizeUsed += TmpPathLen;

        // PDO out length for this module (to assign the length to the pdo configurations)
        pCfg^$USINT := pHelpModule^.ModuleInfo.PdoOutLen;
        pCfg              += sizeof(USINT);
        ConfigMemSizeUsed += sizeof(USINT);

        pHelpModule := pHelpModule^.pNext;
      end_while;

      pCfg := CheckConfigMemSize(sizeof(USINT));
      if pCfg = NIL then
        // error message already logged by function
        return;
      end_if;

      // add number of pdo configurations to memory
      pCfg^$USINT := PdoCfgNo;
      pCfg              += sizeof(USINT);
      ConfigMemSizeUsed += sizeof(USINT);

      // add all pdo configurations to memory (module configs must be available, to find out the PDO length)
      if pFirstPdoCfg then
        pHelpPdo := pFirstPdoCfg;
        // go through list
        while pHelpPdo do
          // add the elements

          // check if we have enough memory to add the next module
          AddConfigSize := sizeof(USINT) + sizeof(BSINT) + sizeof(HDINT) + sizeof(UINT) + pHelpPdo^.PdoInfo.SourcePathLen + sizeof(UINT) + pHelpPdo^.PdoInfo.DestPathLen;
          pCfg := CheckConfigMemSize(AddConfigSize);
          if pCfg = NIL then
            // error message already logged by function
            return;
          end_if;

          // first of all we have to find out the pdo length of this element => search the module configurations until we find our source and copy the pdo length
          if pHelpPdo^.PdoInfo.PdoLen = 0 then
            pHelpModule := pFirstModuleCfg;
            // go through list
            while pHelpModule do
              // if the path of the source module matches, save the pdolength of this module
              if (pHelpPdo^.PdoInfo.SourcePathLen = pHelpModule^.ModuleInfo.PathLen) & (To_StdLib.MemCmp(dest:= pHelpPdo^.PdoInfo.pSourcePath, source:= pHelpModule^.ModuleInfo.pPath , size:= pHelpPdo^.PdoInfo.SourcePathLen) = 0) then
                pHelpPdo^.PdoInfo.PdoLen := pHelpModule^.ModuleInfo.PdoOutLen;
                exit;
              end_if;
              pHelpModule := pHelpModule^.pNext;
            end_while;
          end_if;

          // PDO Length
          pCfg^$USINT := pHelpPdo^.PdoInfo.PdoLen;
          pCfg              += sizeof(USINT);
          ConfigMemSizeUsed += sizeof(USINT);

          // info
          pCfg^$BSINT := pHelpPdo^.PdoInfo.Info;
          pCfg              += sizeof(BSINT);
          ConfigMemSizeUsed += sizeof(BSINT);

          // interface CRC
          pCfg^$HDINT := pHelpPdo^.PdoInfo.InterfaceCRC;
          pCfg              += sizeof(HDINT);
          ConfigMemSizeUsed += sizeof(HDINT);

          // Source Path Length
          TmpPathLen := pHelpPdo^.PdoInfo.SourcePathLen; // save some time with this local variable
          pCfg^$UINT := TmpPathLen;
          pCfg              += sizeof(UINT);
          ConfigMemSizeUsed += sizeof(UINT);

          // Source Path
          _memcpy(ptr1:=pCfg, ptr2:=pHelpPdo^.PdoInfo.pSourcePath, cntr:=TmpPathLen);
          pCfg += TmpPathLen;
          ConfigMemSizeUsed += TmpPathLen;

          // Destination Path Length
          TmpPathLen := pHelpPdo^.PdoInfo.DestPathLen; // save some time with this local variable
          pCfg^$UINT := TmpPathLen;
          pCfg              += sizeof(UINT);
          ConfigMemSizeUsed += sizeof(UINT);

          // Destination Path
          _memcpy(ptr1:=pCfg, ptr2:=pHelpPdo^.PdoInfo.pDestPath, cntr:=TmpPathLen);
          pCfg += TmpPathLen;
          ConfigMemSizeUsed += TmpPathLen;

          pHelpPdo := pHelpPdo^.pNext;
        end_while;
      end_if;

      pCfg := CheckConfigMemSize(sizeof(USINT));
      if pCfg = NIL then
        // error message already logged by function
        return;
      end_if;

      // add number of slave configurations to memory
      pCfg^$USINT       := SlaveCfgNo;
      pCfg              += sizeof(USINT);
      ConfigMemSizeUsed += sizeof(USINT);

      pHelpSlave := pFirstSlaveCfg;
      // go through list
      while pHelpSlave do
        // add the elements

        // check if we have enough memory to add the next module
        AddConfigSize := sizeof(BSINT) + sizeof(HDINT) + sizeof(UINT) + pHelpSlave^.SlaveInfo.PathLen + sizeof(UINT) + pHelpSlave^.SlaveInfo.CompPathLen;

        pCfg := CheckConfigMemSize(AddConfigSize);
        if pCfg = NIL then
          // error message already logged by function
          return;
        end_if;

        // info
        pCfg^$BSINT := pHelpSlave^.SlaveInfo.Info;
        pCfg              += sizeof(BSINT);
        ConfigMemSizeUsed += sizeof(BSINT);

        // InterfaceCRC
        pCfg^$HDINT := pHelpSlave^.SlaveInfo.InterfaceCRC;
        pCfg              += sizeof(HDINT);
        ConfigMemSizeUsed += sizeof(HDINT);

        // uncompressed Slave path
        TmpPathLen := pHelpSlave^.SlaveInfo.PathLen; // save some time with this local variable
        pCfg^$UINT := TmpPathLen;
        pCfg              += sizeof(UINT);
        ConfigMemSizeUsed += sizeof(UINT);

        _memcpy(ptr1:=pCfg, ptr2:=pHelpSlave^.SlaveInfo.pPath, cntr:=TmpPathLen);
        pCfg += TmpPathLen;
        ConfigMemSizeUsed += TmpPathLen;

        // compressed Slave path
        TmpPathLen := pHelpSlave^.SlaveInfo.CompPathLen; // save some time with this local variable
        pCfg^$UINT := TmpPathLen;
        pCfg              += sizeof(UINT);
        ConfigMemSizeUsed += sizeof(UINT);

        _memcpy(ptr1:=pCfg, ptr2:=pHelpSlave^.SlaveInfo.pCompPath, cntr:=TmpPathLen);
        pCfg += TmpPathLen;
        ConfigMemSizeUsed += TmpPathLen;

        pHelpSlave := pHelpSlave^.pNext;
      end_while;

    else
      // add number of module, pdo and slave configurations to memory (all as 0)

      // no module configs
      pCfg^$USINT := 0;
      pCfg              += sizeof(USINT);
      ConfigMemSizeUsed += sizeof(USINT);

      // no pdo configs
      pCfg^$USINT := 0;
      pCfg              += sizeof(USINT);
      ConfigMemSizeUsed += sizeof(USINT);

      // no slave configs
      pCfg^$USINT := 0;
      pCfg              += sizeof(USINT);
      ConfigMemSizeUsed += sizeof(USINT);
    end_if;

    MyPara.uiCmd := CMD_SM_CPU_CFG_TO_MANAGER;
    MyPara.aPara[0] := ConfigMemSizeUsed$DINT;
    MyPara.aPara[1] := pConfigMem$DINT;
    if pSafetyManagerThis^.NewInst(#MyPara, #MyResult) = READY then
      // the manager takes care of our memory from now on
      pFirstSlaveCfg := NIL;
    end_if;

    // now tell the manager, what kind of configuration we have
    MyPara.uiCmd := CMD_SM_NEW_CFG_TYPE;
    MyPara.aPara[0] := SafetyNumber$DINT;
    MyPara.aPara[1] := NewConfigType;
    pSafetyManagerThis^.NewInst(#MyPara, #MyResult);
  else
    LogError("@ZZZZ (SafetyCDIAS_Base::CreateAndSendCfg) No config memory or invalid memory size usage");
  end_if;

END_FUNCTION

#pragma warning(disable: 73)
FUNCTION VIRTUAL SafetyCDIAS_Base::CheckVariant
	VAR_INPUT
		us_ActVariant 	: USINT;
	END_VAR
	VAR_OUTPUT
		b_IsOK 	        : BOOL;
	END_VAR

  // if the overwritten methods are getting deleted, we already have a code for compatiblity here
  b_IsOK := TRUE; // FALSE;

END_FUNCTION
#pragma warning(default: 73)

FUNCTION SafetyCDIAS_Base::SendAllUnsafeValues
  VAR
  	pHelpUnsafeOut : ^UnsafeIORoutingElement;
  END_VAR

  // mark all unsafe values as not sent
  pHelpUnsafeOut := p_UnsafeInputsTable;
  while pHelpUnsafeOut do
    pHelpUnsafeOut^.b_AlreadyTransmitted := FALSE;

    pHelpUnsafeOut := pHelpUnsafeOut^.pNext;
  end_while;

  // reset the actual pointer
  pUnsafeInElement := NIL;

END_FUNCTION

FUNCTION SafetyCDIAS_Base::GetDestinationCRCs
  VAR
    pHelpModule : ^t_ModuleListElem;
    pHelpPdo    : ^t_PdoListElem;
  END_VAR

  // go through the module list
  pHelpModule := pFirstModuleCfg;
  while pHelpModule do
    pHelpPdo := pFirstPdoCfg;
    while pHelpPdo do
      // search in the PDOs if this module is an interface frame destination somewhere
      if pHelpPdo^.PdoInfo.Info.IsInterfacePDO then
        if (pHelpPdo^.PdoInfo.DestPathLen = pHelpModule^.ModuleInfo.PathLen) &
         (To_StdLib.MemCmp(dest:= pHelpModule^.ModuleInfo.pPath, source:= pHelpPdo^.PdoInfo.pDestPath , size:= pHelpModule^.ModuleInfo.PathLen) = 0) then
          pHelpModule^.ModuleInfo.Info.IsInterfaceDest := TRUE;
          if pHelpModule^.ModuleInfo.DestCRCNo & pHelpModule^.ModuleInfo.pDestCRCs then
            pHelpModule^.ModuleInfo.pDestCRCs$^void := To_StdLib.ReAlloc(mptr:=pHelpModule^.ModuleInfo.pDestCRCs, newsize:=(pHelpModule^.ModuleInfo.DestCRCNo+1) * sizeof(HDINT));
          else
            pHelpModule^.ModuleInfo.pDestCRCs$^void := To_StdLib.Malloc(sizeof(HDINT));
          end_if;

          (pHelpModule^.ModuleInfo.pDestCRCs + pHelpModule^.ModuleInfo.DestCRCNo * sizeof(HDINT))^ := pHelpPdo^.PdoInfo.InterfaceCRC;

          pHelpModule^.ModuleInfo.DestCRCNo += 1;
        end_if;
      else
        // if this is module is optional and it's the source of the PDO => the pdo is also optional
        if pHelpModule^.ModuleInfo.Info.IsOptional & (pHelpPdo^.PdoInfo.SourcePathLen = pHelpModule^.ModuleInfo.PathLen) &
         (To_StdLib.MemCmp(dest:= pHelpModule^.ModuleInfo.pPath, source:= pHelpPdo^.PdoInfo.pSourcePath , size:= pHelpModule^.ModuleInfo.PathLen) = 0) then
          pHelpPdo^.PdoInfo.Info.IsOptional := TRUE;
        end_if;
      end_if;

      pHelpPdo := pHelpPdo^.pNext;
    end_while;

    pHelpModule := pHelpModule^.pNext;
  end_while;

END_FUNCTION

FUNCTION SafetyCDIAS_Base::CountBits
	VAR_INPUT
		BitMask 	: BDINT;
	END_VAR
	VAR_OUTPUT
		BitNo 	  : UDINT;
	END_VAR

  BitNo := 0;

  while BitMask do
    BitMask := BitMask AND (BitMask - 1);
    BitNo += 1;
  end_while;

END_FUNCTION

FUNCTION VIRTUAL SafetyCDIAS_Base::IsOptimizedCPU
	VAR_OUTPUT
		IsOptimized 	: DINT;
	END_VAR

  if us_Variant = CSCP012_SERIES then
    IsOptimized := TRUE;
  else
    IsOptimized := FALSE;
  end_if;

END_FUNCTION

FUNCTION VIRTUAL SafetyCDIAS_Base::CheckConfigMemSize
	VAR_INPUT
		AddConfigSize 	: UDINT;
	END_VAR
	VAR_OUTPUT
		pCfg 	          : ^void;
	END_VAR
  VAR
  	pTempMem        : ^void;
  END_VAR

  pCfg := NIL;

  if ((ConfigMemSizeUsed + AddConfigSize) > ConfigMemSize) & (AddConfigSize <= CONFIG_MEMORY_BLOCK_SIZE) then
    // if there isn't enough memory => reallocate
    pTempMem := To_StdLib.ReAlloc(mptr:=pConfigMem, newsize:=ConfigMemSize + CONFIG_MEMORY_BLOCK_SIZE);
    IF pTempMem <> NIL THEN
      pConfigMem := pTempMem;
      ConfigMemSize += CONFIG_MEMORY_BLOCK_SIZE;
    ELSE
      ClassState := _MemAllocFailed;
      LogError("@ZZZZ (SafetyCDIAS_Base::CheckConfigMemSize) Failed to reallocate configuration memory!");
      return;
    END_IF;
  elsif (AddConfigSize > CONFIG_MEMORY_BLOCK_SIZE) then
    ClassState := _MemAllocFailed;
    LogError("@ZZZZ (SafetyCDIAS_Base::CheckConfigMemSize) The configuration of a single config element is too big to handle!");
    return;
  end_if;

  pCfg := pConfigMem + ConfigMemSizeUsed;

END_FUNCTION

FUNCTION SafetyCDIAS_Base::DToH
	VAR_INPUT
		pt 	    : ^CHAR;
		value 	: DINT;
	END_VAR
  VAR
    val     : UDINT;
  END_VAR

  // this method converts a single byte into a zero-terminated hexstring like 0xA4 => "A4"
  val := value$UDINT;

  // zero termination
  (pt + 2)^ := 0;

  // start with the low nibble
  if (val AND 16#F) < 10 then
    (pt + 1)^ := (val AND 16#F)$USINT + '0';
  else
    (pt + 1)^ := (val AND 16#F)$USINT - 10 + 'A';
  end_if;

  // now get the high nibble
  val := val / 16;

  if (val AND 16#F) < 10 then
    pt^ := (val AND 16#F)$USINT + '0';
  else
    pt^ := (val AND 16#F)$USINT - 10 + 'A';
  end_if;

END_FUNCTION

FUNCTION SafetyCDIAS_Base::LogHWPath
	VAR_INPUT
		pString 	: ^CHAR;
		pHWPath 	: ^USINT;
	END_VAR
  VAR
    TempStr   : ARRAY [0..99] OF CHAR;
    TraceVal  : USINT;
    i         : UINT;
    MyMsg     : ARRAY [0..599] OF CHAR;
  END_VAR

  if pString & pHWPath then

    _strncpy(dest:=#MyMsg[0], src:=pString, max:=200);

    TraceVal := pHWPath^;
    if TraceVal then
      TraceVal  += 2; //show also the length
      i         := 0;
      while (TraceVal >= 1) & (i < 95) do
        DToH(#TempStr[i], pHWPath^$USINT);
        i         += 2; // 2 chars per byte
        TempStr[i]:= ' ';
        i         += 1;
        pHWPath   += 1;
        TraceVal  -= 1;
      end_while;
      TempStr[i] := 0;

      _strcat( dest:=#MyMsg[0], src:=#TempStr[0]);
    end_if;

#ifdef HWC_LogError
    HWC_LogError(this, #MyMsg[0]);
#endif
  end_if;

END_FUNCTION

FUNCTION VIRTUAL GLOBAL SafetyCDIAS_Base::QuitComError::Write
	VAR_INPUT
		input (EAX) 	: DINT;
	END_VAR
	VAR_OUTPUT
		result (EAX) 	: DINT;
	END_VAR

 	result := input;

  if b_QuitErrorAvailable then
    // remember to do it in next background
    QuitComError := 2;
  else
    // remember. that there has been a manual quit (for writing PDOs in PostScan)
    b_ManualQuit := TRUE;

    // remember to do it in next cyclic
    QuitComError := 1;
  end_if;

END_FUNCTION

FUNCTION VIRTUAL SafetyCDIAS_Base::GetFWVersion
	VAR_INPUT
		pData 	: ^CHAR;
		length 	: DINT;
	END_VAR

  //Check pointer
  if pData then
    //Length of Firmwareversion (HDINT) -> 8Byte +1 byte zero termination
    if Length >= 9 then
      _itoa(udNumber:=FW_Version, pString:=pData);
    else
      pData^ := 0;
    end_if;
  end_if;

END_FUNCTION

FUNCTION VIRTUAL GLOBAL SafetyCDIAS_Base::GetDiagConnect::NewInst
	VAR_INPUT
		pPara 	  : ^CmdStruct;
		pResult 	: ^Results;
	END_VAR
	VAR_OUTPUT
		ret_code 	: IprStates;
	END_VAR
